(* IEC 61131-3 sources: plc-st-coding-agent/progress/evidence/f14_v10_full_20261113/jobs/custom_deepseek-v4pro (part 2) *)

(* ---- public-hard-02.raw_candidate_04.st ---- *)
(* ENGINEERING_CONTRACT
- Outputs conveyorLeft/deactivate in IDLE, PROCESSING and DONE; active only in MOVING state; no latch. PUB005.
- State machine: 0=IDLE waits sensor1 AND station1Start with valid length; 1=MOVING waits arrival at target sensor; 2=PROCESSING waits completion at current station 2..4; 3=DONE after station 5 arrival. PUB001/PUB002/PUB005.
- Movement direction: target station > current -> conveyorRight; target < current -> conveyorLeft; target == current stays at station for repeated processing step. PUB005.
- Completion signals are level-sensitive; on receiving completion, step advances, next sequence entry is queried, and movement restarts toward that station. PUB002.
- Final active sequence entry is station 5; arrival at 5 stops conveyor and enters DONE. A new start is permitted from DONE when the start condition is true. PUB003/PUB006.
- processLength validated 1..8; dynamic array indexing bounded by processLength; sequence values assumed to satisfy contract (2..4 processing, final 5). PUB004.
- Unspecified: exact restart behavior after DONE is level-sensitive on sensor1 and station1Start. No explicit reset input is used.
*)
(* CONTRACT_RULES [] *)
FUNCTION_BLOCK FlexibleProcessingControl
VAR_INPUT
    processLength : USINT;
    sensor1 : BOOL;
    sensor2 : BOOL;
    sensor3 : BOOL;
    sensor4 : BOOL;
    sensor5 : BOOL;
    station1Start : BOOL;
    station2Complete : BOOL;
    station3Complete : BOOL;
    station4Complete : BOOL;
    processSequence : ARRAY[1..8] OF USINT;
END_VAR
VAR_OUTPUT
    conveyorLeft : BOOL;
    conveyorRight : BOOL;
END_VAR
VAR
    local_state : USINT := 0; (* 0 = idle, 1 = moving, 2 = processing, 3 = done *)
    local_step : USINT := 0;
    local_target : USINT := 0;
    local_currentStation : USINT := 1;
    local_moveLeft : BOOL := FALSE;
    local_moveRight : BOOL := FALSE;
    local_arrival : BOOL := FALSE;
    local_complete : BOOL := FALSE;
END_VAR

(* Default outputs deactivated unless set by MOVING state *)
conveyorLeft := FALSE;
conveyorRight := FALSE;

CASE local_state OF
0: (* IDLE: wait for raw material at station 1 and start button *)
    IF processLength >= 1 AND processLength <= 8 AND sensor1 AND station1Start THEN
        local_step := 1;
        local_target := processSequence[1];
        local_currentStation := 1;
        IF local_target > local_currentStation THEN
            local_moveLeft := FALSE;
            local_moveRight := TRUE;
            conveyorLeft := FALSE;
            conveyorRight := TRUE;
            local_state := 1;
        ELSIF local_target < local_currentStation THEN
            local_moveLeft := TRUE;
            local_moveRight := FALSE;
            conveyorLeft := TRUE;
            conveyorRight := FALSE;
            local_state := 1;
        END_IF;
    END_IF;

1: (* MOVING: drive conveyor in chosen direction until target sensor detects arrival *)
    conveyorLeft := local_moveLeft;
    conveyorRight := local_moveRight;

    local_arrival := FALSE;
    IF local_target = 1 AND sensor1 THEN
        local_arrival := TRUE;
    ELSIF local_target = 2 AND sensor2 THEN
        local_arrival := TRUE;
    ELSIF local_target = 3 AND sensor3 THEN
        local_arrival := TRUE;
    ELSIF local_target = 4 AND sensor4 THEN
        local_arrival := TRUE;
    ELSIF local_target = 5 AND sensor5 THEN
        local_arrival := TRUE;
    END_IF;

    IF local_arrival THEN
        conveyorLeft := FALSE;
        conveyorRight := FALSE;
        local_moveLeft := FALSE;
        local_moveRight := FALSE;
        local_currentStation := local_target;

        IF local_currentStation = 5 THEN
            local_state := 3; (* final output station reached *)
        ELSE
            local_state := 2; (* processing station reached *)
        END_IF;
    END_IF;

2: (* PROCESSING: wait for completion signal at current processing station *)
    local_complete := FALSE;
    IF local_currentStation = 2 THEN
        local_complete := station2Complete;
    ELSIF local_currentStation = 3 THEN
        local_complete := station3Complete;
    ELSIF local_currentStation = 4 THEN
        local_complete := station4Complete;
    END_IF;

    IF local_complete THEN
        IF local_step < processLength THEN
            local_step := local_step + 1;
            local_target := processSequence[local_step];

            IF local_target > local_currentStation THEN
                local_moveLeft := FALSE;
                local_moveRight := TRUE;
                conveyorLeft := FALSE;
                conveyorRight := TRUE;
                local_state := 1;
            ELSIF local_target < local_currentStation THEN
                local_moveLeft := TRUE;
                local_moveRight := FALSE;
                conveyorLeft := TRUE;
                conveyorRight := FALSE;
                local_state := 1;
            ELSE
                (* Same station: remain in processing for the next sequence entry *)
                local_state := 2;
            END_IF;
        ELSE
            (* Invalid sequence: current processing station is not followed by final station 5 *)
            local_state := 3;
        END_IF;
    END_IF;

3: (* DONE: product delivered to station 5; optionally wait for next start *)
    IF processLength >= 1 AND processLength <= 8 AND sensor1 AND station1Start THEN
        local_step := 1;
        local_target := processSequence[1];
        local_currentStation := 1;
        IF local_target > local_currentStation THEN
            local_moveLeft := FALSE;
            local_moveRight := TRUE;
            conveyorLeft := FALSE;
            conveyorRight := TRUE;
            local_state := 1;
        ELSIF local_target < local_currentStation THEN
            local_moveLeft := TRUE;
            local_moveRight := FALSE;
            conveyorLeft := TRUE;
            conveyorRight := FALSE;
            local_state := 1;
        END_IF;
    END_IF;
END_CASE;

END_FUNCTION_BLOCK

(* ---- public-hard-03.candidate_01.st ---- *)
TYPE ST_Recipe :
STRUCT
    recipeID : INT;
    ingredientType : INT;
    ingredientRatio : REAL;
    productionTemperature : REAL;
END_STRUCT
END_TYPE;

FUNCTION_BLOCK FB_RecipeManagement
VAR_INPUT
    addRecipe : BOOL;
    deleteRecipe : BOOL;
    modifyRecipe : BOOL;
    queryRecipe : BOOL;
    recipeIn : ST_Recipe;
END_VAR
VAR_OUTPUT
    recipeAdded : BOOL;
    recipeDeleted : BOOL;
    recipeModified : BOOL;
    recipeQueryResult : ST_Recipe;
    error : BOOL;
    status : WORD;
END_VAR
VAR_IN_OUT
    recipe : ARRAY[1..10] OF ST_Recipe;
END_VAR
VAR
    tmp_i : INT;
    tmp_found : BOOL;
    tmp_index : INT;
    tmp_emptyIndex : INT;
    tmp_cmdCount : INT;
    tmp_emptyRecipe : ST_Recipe;
END_VAR

(*
ENGINEERING_CONTRACT
recipeAdded/Deleted/Modified: pulse TRUE only when exactly one matching request is TRUE and operation succeeds; not latched.
recipeQueryResult: valid only on successful query; otherwise zero struct. Not latched.
error/status: same-scan result; success/no command => error=FALSE,status=0. Error codes PUB003-PUB005, multiple commands => 16#8006.
recipe IN_OUT: caller retains; changed only on successful add/delete/modify. Add uses smallest empty index (PUB003).
Search ignores slots where recipeID=0. Units: raw REAL values; no scaling. Simultaneous commands are unsupported and modify nothing.
*)

(* CONTRACT_RULES [] *)

tmp_emptyRecipe.recipeID := 0;
tmp_emptyRecipe.ingredientType := 0;
tmp_emptyRecipe.ingredientRatio := 0.0;
tmp_emptyRecipe.productionTemperature := 0.0;

recipeAdded := FALSE;
recipeDeleted := FALSE;
recipeModified := FALSE;
recipeQueryResult := tmp_emptyRecipe;
error := FALSE;
status := 0;

tmp_cmdCount := 0;
IF addRecipe THEN
    tmp_cmdCount := tmp_cmdCount + 1;
END_IF;
IF deleteRecipe THEN
    tmp_cmdCount := tmp_cmdCount + 1;
END_IF;
IF modifyRecipe THEN
    tmp_cmdCount := tmp_cmdCount + 1;
END_IF;
IF queryRecipe THEN
    tmp_cmdCount := tmp_cmdCount + 1;
END_IF;

IF tmp_cmdCount > 1 THEN
    error := TRUE;
    status := 16#8006;
    RETURN;
END_IF;

IF addRecipe THEN
    tmp_found := FALSE;
    tmp_index := 0;
    FOR tmp_i := 1 TO 10 DO
        IF (recipe[tmp_i].recipeID <> 0) AND (recipe[tmp_i].recipeID = recipeIn.recipeID) THEN
            tmp_found := TRUE;
            tmp_index := tmp_i;
            EXIT;
        END_IF;
    END_FOR;

    IF tmp_found THEN
        error := TRUE;
        status := 16#8002;
    ELSE
        tmp_emptyIndex := 0;
        FOR tmp_i := 1 TO 10 DO
            IF recipe[tmp_i].recipeID = 0 THEN
                tmp_emptyIndex := tmp_i;
                EXIT;
            END_IF;
        END_FOR;

        IF tmp_emptyIndex = 0 THEN
            error := TRUE;
            status := 16#8003;
        ELSE
            recipe[tmp_emptyIndex] := recipeIn;
            recipeAdded := TRUE;
            error := FALSE;
            status := 0;
        END_IF;
    END_IF;
END_IF;

IF deleteRecipe THEN
    tmp_found := FALSE;
    tmp_index := 0;
    FOR tmp_i := 1 TO 10 DO
        IF (recipe[tmp_i].recipeID <> 0) AND (recipe[tmp_i].recipeID = recipeIn.recipeID) THEN
            tmp_found := TRUE;
            tmp_index := tmp_i;
            EXIT;
        END_IF;
    END_FOR;

    IF NOT tmp_found THEN
        error := TRUE;
        status := 16#8004;
    ELSE
        recipe[tmp_index] := tmp_emptyRecipe;
        recipeDeleted := TRUE;
        error := FALSE;
        status := 0;
    END_IF;
END_IF;

IF modifyRecipe THEN
    tmp_found := FALSE;
    tmp_index := 0;
    FOR tmp_i := 1 TO 10 DO
        IF (recipe[tmp_i].recipeID <> 0) AND (recipe[tmp_i].recipeID = recipeIn.recipeID) THEN
            tmp_found := TRUE;
            tmp_index := tmp_i;
            EXIT;
        END_IF;
    END_FOR;

    IF NOT tmp_found THEN
        error := TRUE;
        status := 16#8005;
    ELSE
        recipe[tmp_index] := recipeIn;
        recipeModified := TRUE;
        error := FALSE;
        status := 0;
    END_IF;
END_IF;

IF queryRecipe THEN
    tmp_found := FALSE;
    tmp_index := 0;
    FOR tmp_i := 1 TO 10 DO
        IF (recipe[tmp_i].recipeID <> 0) AND (recipe[tmp_i].recipeID = recipeIn.recipeID) THEN
            tmp_found := TRUE;
            tmp_index := tmp_i;
            EXIT;
        END_IF;
    END_FOR;

    IF NOT tmp_found THEN
        error := TRUE;
        status := 16#8001;
    ELSE
        recipeQueryResult := recipe[tmp_index];
        error := FALSE;
        status := 0;
    END_IF;
END_IF;

END_FUNCTION_BLOCK

(* ---- public-hard-03.candidate_02.st ---- *)
TYPE ST_Recipe :
STRUCT
    recipeID : INT;
    ingredientType : INT;
    ingredientRatio : REAL;
    productionTemperature : REAL;
END_STRUCT
END_TYPE;

FUNCTION_BLOCK FB_RecipeManagement
VAR_INPUT
    addRecipe : BOOL;
    deleteRecipe : BOOL;
    modifyRecipe : BOOL;
    queryRecipe : BOOL;
    recipeIn : ST_Recipe;
END_VAR
VAR_OUTPUT
    recipeAdded : BOOL;
    recipeDeleted : BOOL;
    recipeModified : BOOL;
    recipeQueryResult : ST_Recipe;
    error : BOOL;
    status : WORD;
END_VAR
VAR_IN_OUT
    recipe : ARRAY[1..10] OF ST_Recipe;
END_VAR
VAR
    tmp_i : INT;
    tmp_found : BOOL;
    tmp_index : INT;
    tmp_emptyIndex : INT;
    tmp_cmdCount : INT;
    tmp_emptyRecipe : ST_Recipe;
    tmp_addReq : BOOL;
    tmp_deleteReq : BOOL;
    tmp_modifyReq : BOOL;
    tmp_queryReq : BOOL;
    prevAdd : BOOL := FALSE;
    prevDelete : BOOL := FALSE;
    prevModify : BOOL := FALSE;
    prevQuery : BOOL := FALSE;
END_VAR

(*
ENGINEERING_CONTRACT
Request signals are edge-triggered (rising edge only).
recipeAdded/Deleted/Modified: one-scan pulse on successful operation; otherwise FALSE.
recipeQueryResult: valid only in the scan of a successful query; zero struct otherwise.
error/status: same-scan result; success/no edge => error=FALSE,status=0.
Simultaneous rising command edges => error=TRUE,status=16#8006; database unchanged.
Database in recipe[] retains state between scans; add uses smallest empty index.
*)

(* CONTRACT_RULES [] *)

tmp_emptyRecipe.recipeID := 0;
tmp_emptyRecipe.ingredientType := 0;
tmp_emptyRecipe.ingredientRatio := 0.0;
tmp_emptyRecipe.productionTemperature := 0.0;

recipeAdded := FALSE;
recipeDeleted := FALSE;
recipeModified := FALSE;
recipeQueryResult := tmp_emptyRecipe;
error := FALSE;
status := 0;

tmp_addReq := addRecipe AND NOT prevAdd;
tmp_deleteReq := deleteRecipe AND NOT prevDelete;
tmp_modifyReq := modifyRecipe AND NOT prevModify;
tmp_queryReq := queryRecipe AND NOT prevQuery;

prevAdd := addRecipe;
prevDelete := deleteRecipe;
prevModify := modifyRecipe;
prevQuery := queryRecipe;

tmp_cmdCount := 0;
IF tmp_addReq THEN
    tmp_cmdCount := tmp_cmdCount + 1;
END_IF;
IF tmp_deleteReq THEN
    tmp_cmdCount := tmp_cmdCount + 1;
END_IF;
IF tmp_modifyReq THEN
    tmp_cmdCount := tmp_cmdCount + 1;
END_IF;
IF tmp_queryReq THEN
    tmp_cmdCount := tmp_cmdCount + 1;
END_IF;

IF tmp_cmdCount > 1 THEN
    error := TRUE;
    status := 16#8006;
    RETURN;
END_IF;

IF tmp_addReq THEN
    tmp_found := FALSE;
    tmp_index := 0;
    FOR tmp_i := 1 TO 10 DO
        IF (recipe[tmp_i].recipeID <> 0) AND (recipe[tmp_i].recipeID = recipeIn.recipeID) THEN
            tmp_found := TRUE;
            tmp_index := tmp_i;
            EXIT;
        END_IF;
    END_FOR;

    IF tmp_found THEN
        error := TRUE;
        status := 16#8002;
    ELSE
        tmp_emptyIndex := 0;
        FOR tmp_i := 1 TO 10 DO
            IF recipe[tmp_i].recipeID = 0 THEN
                tmp_emptyIndex := tmp_i;
                EXIT;
            END_IF;
        END_FOR;

        IF tmp_emptyIndex = 0 THEN
            error := TRUE;
            status := 16#8003;
        ELSE
            recipe[tmp_emptyIndex] := recipeIn;
            recipeAdded := TRUE;
            error := FALSE;
            status := 0;
        END_IF;
    END_IF;
END_IF;

IF tmp_deleteReq THEN
    tmp_found := FALSE;
    tmp_index := 0;
    FOR tmp_i := 1 TO 10 DO
        IF (recipe[tmp_i].recipeID <> 0) AND (recipe[tmp_i].recipeID = recipeIn.recipeID) THEN
            tmp_found := TRUE;
            tmp_index := tmp_i;
            EXIT;
        END_IF;
    END_FOR;

    IF NOT tmp_found THEN
        error := TRUE;
        status := 16#8004;
    ELSE
        recipe[tmp_index] := tmp_emptyRecipe;
        recipeDeleted := TRUE;
        error := FALSE;
        status := 0;
    END_IF;
END_IF;

IF tmp_modifyReq THEN
    tmp_found := FALSE;
    tmp_index := 0;
    FOR tmp_i := 1 TO 10 DO
        IF (recipe[tmp_i].recipeID <> 0) AND (recipe[tmp_i].recipeID = recipeIn.recipeID) THEN
            tmp_found := TRUE;
            tmp_index := tmp_i;
            EXIT;
        END_IF;
    END_FOR;

    IF NOT tmp_found THEN
        error := TRUE;
        status := 16#8005;
    ELSE
        recipe[tmp_index] := recipeIn;
        recipeModified := TRUE;
        error := FALSE;
        status := 0;
    END_IF;
END_IF;

IF tmp_queryReq THEN
    tmp_found := FALSE;
    tmp_index := 0;
    FOR tmp_i := 1 TO 10 DO
        IF (recipe[tmp_i].recipeID <> 0) AND (recipe[tmp_i].recipeID = recipeIn.recipeID) THEN
            tmp_found := TRUE;
            tmp_index := tmp_i;
            EXIT;
        END_IF;
    END_FOR;

    IF NOT tmp_found THEN
        error := TRUE;
        status := 16#8001;
    ELSE
        recipeQueryResult := recipe[tmp_index];
        error := FALSE;
        status := 0;
    END_IF;
END_IF;

END_FUNCTION_BLOCK

(* ---- public-hard-03.candidate_03.st ---- *)
TYPE ST_Recipe :
STRUCT
    recipeID : INT;
    ingredientType : INT;
    ingredientRatio : REAL;
    productionTemperature : REAL;
END_STRUCT
END_TYPE;

FUNCTION_BLOCK FB_RecipeManagement
VAR_INPUT
    addRecipe : BOOL;
    deleteRecipe : BOOL;
    modifyRecipe : BOOL;
    queryRecipe : BOOL;
    recipeIn : ST_Recipe;
END_VAR
VAR_OUTPUT
    recipeAdded : BOOL;
    recipeDeleted : BOOL;
    recipeModified : BOOL;
    recipeQueryResult : ST_Recipe;
    error : BOOL;
    status : WORD;
END_VAR
VAR_IN_OUT
    recipe : ARRAY[1..10] OF ST_Recipe;
END_VAR
VAR
    tmp_i : INT;
    tmp_found : BOOL;
    tmp_index : INT;
    tmp_emptyIndex : INT;
    tmp_emptyRecipe : ST_Recipe;
END_VAR

(*
ENGINEERING_CONTRACT
recipeAdded/Deleted/Modified: pulse TRUE only when corresponding request is TRUE and operation succeeds; not latched.
recipeQueryResult: valid only on successful query; otherwise zero struct. Not latched.
error/status: same-scan result; success/no command => error=FALSE,status=0.
Search ignores slots where recipeID=0. Units: raw REAL values; no scaling.
Simultaneous commands are not specified by the public contract; implementation processes all active commands in the
present scan using the defined operation order add, delete, modify, query. No extra priority or 8006 code is invented.
*)

(* CONTRACT_RULES [] *)

tmp_emptyRecipe.recipeID := 0;
tmp_emptyRecipe.ingredientType := 0;
tmp_emptyRecipe.ingredientRatio := 0.0;
tmp_emptyRecipe.productionTemperature := 0.0;

recipeAdded := FALSE;
recipeDeleted := FALSE;
recipeModified := FALSE;
recipeQueryResult := tmp_emptyRecipe;
error := FALSE;
status := 0;

IF addRecipe THEN
    tmp_found := FALSE;
    tmp_index := 0;
    FOR tmp_i := 1 TO 10 DO
        IF (recipe[tmp_i].recipeID <> 0) AND (recipe[tmp_i].recipeID = recipeIn.recipeID) THEN
            tmp_found := TRUE;
            tmp_index := tmp_i;
            EXIT;
        END_IF;
    END_FOR;

    IF tmp_found THEN
        error := TRUE;
        status := 16#8002;
    ELSE
        tmp_emptyIndex := 0;
        FOR tmp_i := 1 TO 10 DO
            IF recipe[tmp_i].recipeID = 0 THEN
                tmp_emptyIndex := tmp_i;
                EXIT;
            END_IF;
        END_FOR;

        IF tmp_emptyIndex = 0 THEN
            error := TRUE;
            status := 16#8003;
        ELSE
            recipe[tmp_emptyIndex] := recipeIn;
            recipeAdded := TRUE;
            error := FALSE;
            status := 0;
        END_IF;
    END_IF;
END_IF;

IF deleteRecipe THEN
    tmp_found := FALSE;
    tmp_index := 0;
    FOR tmp_i := 1 TO 10 DO
        IF (recipe[tmp_i].recipeID <> 0) AND (recipe[tmp_i].recipeID = recipeIn.recipeID) THEN
            tmp_found := TRUE;
            tmp_index := tmp_i;
            EXIT;
        END_IF;
    END_FOR;

    IF NOT tmp_found THEN
        error := TRUE;
        status := 16#8004;
    ELSE
        recipe[tmp_index] := tmp_emptyRecipe;
        recipeDeleted := TRUE;
        error := FALSE;
        status := 0;
    END_IF;
END_IF;

IF modifyRecipe THEN
    tmp_found := FALSE;
    tmp_index := 0;
    FOR tmp_i := 1 TO 10 DO
        IF (recipe[tmp_i].recipeID <> 0) AND (recipe[tmp_i].recipeID = recipeIn.recipeID) THEN
            tmp_found := TRUE;
            tmp_index := tmp_i;
            EXIT;
        END_IF;
    END_FOR;

    IF NOT tmp_found THEN
        error := TRUE;
        status := 16#8005;
    ELSE
        recipe[tmp_index] := recipeIn;
        recipeModified := TRUE;
        error := FALSE;
        status := 0;
    END_IF;
END_IF;

IF queryRecipe THEN
    tmp_found := FALSE;
    tmp_index := 0;
    FOR tmp_i := 1 TO 10 DO
        IF (recipe[tmp_i].recipeID <> 0) AND (recipe[tmp_i].recipeID = recipeIn.recipeID) THEN
            tmp_found := TRUE;
            tmp_index := tmp_i;
            EXIT;
        END_IF;
    END_FOR;

    IF NOT tmp_found THEN
        error := TRUE;
        status := 16#8001;
    ELSE
        recipeQueryResult := recipe[tmp_index];
        error := FALSE;
        status := 0;
    END_IF;
END_IF;

END_FUNCTION_BLOCK

(* ---- public-hard-03.candidate_04.st ---- *)
TYPE ST_Recipe :
STRUCT
    recipeID : INT;
    ingredientType : INT;
    ingredientRatio : REAL;
    productionTemperature : REAL;
END_STRUCT
END_TYPE;

FUNCTION_BLOCK FB_RecipeManagement
VAR_INPUT
    addRecipe : BOOL;
    deleteRecipe : BOOL;
    modifyRecipe : BOOL;
    queryRecipe : BOOL;
    recipeIn : ST_Recipe;
END_VAR
VAR_OUTPUT
    recipeAdded : BOOL;
    recipeDeleted : BOOL;
    recipeModified : BOOL;
    recipeQueryResult : ST_Recipe;
    error : BOOL;
    status : WORD;
END_VAR
VAR_IN_OUT
    recipe : ARRAY[1..10] OF ST_Recipe;
END_VAR
VAR
    tmp_i : INT;
    tmp_found : BOOL;
    tmp_index : INT;
    tmp_emptyIndex : INT;
    tmp_cmdCount : INT;
    tmp_emptyRecipe : ST_Recipe;
END_VAR

(*
ENGINEERING_CONTRACT
recipeAdded/Deleted/Modified: pulse TRUE only when exactly one matching request is TRUE and operation succeeds; not latched.
recipeQueryResult: valid only on successful query; otherwise zero struct. Not latched.
error/status: same-scan result; success/no command => error=FALSE,status=0. Error codes PUB003-PUB005, multiple commands => 16#8006.
recipe IN_OUT: caller retains; changed only on successful add/delete/modify. Add uses smallest empty index (PUB003).
Search ignores slots where recipeID=0 for query/delete/modify. Add treats recipeIn.recipeID=0 as reserved/invalid and never stores it.
Units: raw REAL values; no scaling. Simultaneous commands are unsupported and modify nothing.
*)

(* CONTRACT_RULES [] *)

tmp_emptyRecipe.recipeID := 0;
tmp_emptyRecipe.ingredientType := 0;
tmp_emptyRecipe.ingredientRatio := 0.0;
tmp_emptyRecipe.productionTemperature := 0.0;

recipeAdded := FALSE;
recipeDeleted := FALSE;
recipeModified := FALSE;
recipeQueryResult := tmp_emptyRecipe;
error := FALSE;
status := 0;

tmp_cmdCount := 0;
IF addRecipe THEN
    tmp_cmdCount := tmp_cmdCount + 1;
END_IF;
IF deleteRecipe THEN
    tmp_cmdCount := tmp_cmdCount + 1;
END_IF;
IF modifyRecipe THEN
    tmp_cmdCount := tmp_cmdCount + 1;
END_IF;
IF queryRecipe THEN
    tmp_cmdCount := tmp_cmdCount + 1;
END_IF;

IF tmp_cmdCount > 1 THEN
    error := TRUE;
    status := 16#8006;
    RETURN;
END_IF;

IF addRecipe THEN
    tmp_found := FALSE;
    tmp_index := 0;
    FOR tmp_i := 1 TO 10 DO
        IF recipe[tmp_i].recipeID = recipeIn.recipeID THEN
            tmp_found := TRUE;
            tmp_index := tmp_i;
            EXIT;
        END_IF;
    END_FOR;

    IF tmp_found THEN
        error := TRUE;
        status := 16#8002;
    ELSE
        tmp_emptyIndex := 0;
        FOR tmp_i := 1 TO 10 DO
            IF recipe[tmp_i].recipeID = 0 THEN
                tmp_emptyIndex := tmp_i;
                EXIT;
            END_IF;
        END_FOR;

        IF tmp_emptyIndex = 0 THEN
            error := TRUE;
            status := 16#8003;
        ELSE
            recipe[tmp_emptyIndex] := recipeIn;
            recipeAdded := TRUE;
            error := FALSE;
            status := 0;
        END_IF;
    END_IF;
END_IF;

IF deleteRecipe THEN
    tmp_found := FALSE;
    tmp_index := 0;
    FOR tmp_i := 1 TO 10 DO
        IF (recipe[tmp_i].recipeID <> 0) AND (recipe[tmp_i].recipeID = recipeIn.recipeID) THEN
            tmp_found := TRUE;
            tmp_index := tmp_i;
            EXIT;
        END_IF;
    END_FOR;

    IF NOT tmp_found THEN
        error := TRUE;
        status := 16#8004;
    ELSE
        recipe[tmp_index] := tmp_emptyRecipe;
        recipeDeleted := TRUE;
        error := FALSE;
        status := 0;
    END_IF;
END_IF;

IF modifyRecipe THEN
    tmp_found := FALSE;
    tmp_index := 0;
    FOR tmp_i := 1 TO 10 DO
        IF (recipe[tmp_i].recipeID <> 0) AND (recipe[tmp_i].recipeID = recipeIn.recipeID) THEN
            tmp_found := TRUE;
            tmp_index := tmp_i;
            EXIT;
        END_IF;
    END_FOR;

    IF NOT tmp_found THEN
        error := TRUE;
        status := 16#8005;
    ELSE
        recipe[tmp_index] := recipeIn;
        recipeModified := TRUE;
        error := FALSE;
        status := 0;
    END_IF;
END_IF;

IF queryRecipe THEN
    tmp_found := FALSE;
    tmp_index := 0;
    FOR tmp_i := 1 TO 10 DO
        IF (recipe[tmp_i].recipeID <> 0) AND (recipe[tmp_i].recipeID = recipeIn.recipeID) THEN
            tmp_found := TRUE;
            tmp_index := tmp_i;
            EXIT;
        END_IF;
    END_FOR;

    IF NOT tmp_found THEN
        error := TRUE;
        status := 16#8001;
    ELSE
        recipeQueryResult := recipe[tmp_index];
        error := FALSE;
        status := 0;
    END_IF;
END_IF;

END_FUNCTION_BLOCK

(* ---- public-hard-03.raw_candidate_01.st ---- *)
TYPE ST_Recipe :
STRUCT
    recipeID : INT;
    ingredientType : INT;
    ingredientRatio : REAL;
    productionTemperature : REAL;
END_STRUCT
END_TYPE

FUNCTION_BLOCK FB_RecipeManagement
VAR_INPUT
    addRecipe : BOOL;
    deleteRecipe : BOOL;
    modifyRecipe : BOOL;
    queryRecipe : BOOL;
    recipeIn : ST_Recipe;
END_VAR
VAR_OUTPUT
    recipeAdded : BOOL;
    recipeDeleted : BOOL;
    recipeModified : BOOL;
    recipeQueryResult : ST_Recipe;
    error : BOOL;
    status : WORD;
END_VAR
VAR_IN_OUT
    recipe : ARRAY[1..10] OF ST_Recipe;
END_VAR
VAR
    tmp_i : INT;
    tmp_found : BOOL;
    tmp_index : INT;
    tmp_emptyIndex : INT;
    tmp_cmdCount : INT;
    tmp_emptyRecipe : ST_Recipe;
END_VAR

(*
ENGINEERING_CONTRACT
recipeAdded/Deleted/Modified: pulse TRUE only when exactly one matching request is TRUE and operation succeeds; not latched.
recipeQueryResult: valid only on successful query; otherwise zero struct. Not latched.
error/status: same-scan result; success/no command => error=FALSE,status=0. Error codes PUB003-PUB005, multiple commands => 16#8006.
recipe IN_OUT: caller retains; changed only on successful add/delete/modify. Add uses smallest empty index (PUB003).
Search ignores slots where recipeID=0. Units: raw REAL values; no scaling. Simultaneous commands are unsupported and modify nothing.
*)

(* CONTRACT_RULES [] *)

tmp_emptyRecipe.recipeID := 0;
tmp_emptyRecipe.ingredientType := 0;
tmp_emptyRecipe.ingredientRatio := 0.0;
tmp_emptyRecipe.productionTemperature := 0.0;

recipeAdded := FALSE;
recipeDeleted := FALSE;
recipeModified := FALSE;
recipeQueryResult := tmp_emptyRecipe;
error := FALSE;
status := 0;

tmp_cmdCount := 0;
IF addRecipe THEN
    tmp_cmdCount := tmp_cmdCount + 1;
END_IF;
IF deleteRecipe THEN
    tmp_cmdCount := tmp_cmdCount + 1;
END_IF;
IF modifyRecipe THEN
    tmp_cmdCount := tmp_cmdCount + 1;
END_IF;
IF queryRecipe THEN
    tmp_cmdCount := tmp_cmdCount + 1;
END_IF;

IF tmp_cmdCount > 1 THEN
    error := TRUE;
    status := 16#8006;
    RETURN;
END_IF;

IF addRecipe THEN
    tmp_found := FALSE;
    tmp_index := 0;
    FOR tmp_i := 1 TO 10 DO
        IF (recipe[tmp_i].recipeID <> 0) AND (recipe[tmp_i].recipeID = recipeIn.recipeID) THEN
            tmp_found := TRUE;
            tmp_index := tmp_i;
            EXIT;
        END_IF;
    END_FOR;

    IF tmp_found THEN
        error := TRUE;
        status := 16#8002;
    ELSE
        tmp_emptyIndex := 0;
        FOR tmp_i := 1 TO 10 DO
            IF recipe[tmp_i].recipeID = 0 THEN
                tmp_emptyIndex := tmp_i;
                EXIT;
            END_IF;
        END_FOR;

        IF tmp_emptyIndex = 0 THEN
            error := TRUE;
            status := 16#8003;
        ELSE
            recipe[tmp_emptyIndex] := recipeIn;
            recipeAdded := TRUE;
            error := FALSE;
            status := 0;
        END_IF;
    END_IF;
END_IF;

IF deleteRecipe THEN
    tmp_found := FALSE;
    tmp_index := 0;
    FOR tmp_i := 1 TO 10 DO
        IF (recipe[tmp_i].recipeID <> 0) AND (recipe[tmp_i].recipeID = recipeIn.recipeID) THEN
            tmp_found := TRUE;
            tmp_index := tmp_i;
            EXIT;
        END_IF;
    END_FOR;

    IF NOT tmp_found THEN
        error := TRUE;
        status := 16#8004;
    ELSE
        recipe[tmp_index] := tmp_emptyRecipe;
        recipeDeleted := TRUE;
        error := FALSE;
        status := 0;
    END_IF;
END_IF;

IF modifyRecipe THEN
    tmp_found := FALSE;
    tmp_index := 0;
    FOR tmp_i := 1 TO 10 DO
        IF (recipe[tmp_i].recipeID <> 0) AND (recipe[tmp_i].recipeID = recipeIn.recipeID) THEN
            tmp_found := TRUE;
            tmp_index := tmp_i;
            EXIT;
        END_IF;
    END_FOR;

    IF NOT tmp_found THEN
        error := TRUE;
        status := 16#8005;
    ELSE
        recipe[tmp_index] := recipeIn;
        recipeModified := TRUE;
        error := FALSE;
        status := 0;
    END_IF;
END_IF;

IF queryRecipe THEN
    tmp_found := FALSE;
    tmp_index := 0;
    FOR tmp_i := 1 TO 10 DO
        IF (recipe[tmp_i].recipeID <> 0) AND (recipe[tmp_i].recipeID = recipeIn.recipeID) THEN
            tmp_found := TRUE;
            tmp_index := tmp_i;
            EXIT;
        END_IF;
    END_FOR;

    IF NOT tmp_found THEN
        error := TRUE;
        status := 16#8001;
    ELSE
        recipeQueryResult := recipe[tmp_index];
        error := FALSE;
        status := 0;
    END_IF;
END_IF;

END_FUNCTION_BLOCK

(* ---- public-hard-03.raw_candidate_02.st ---- *)
TYPE ST_Recipe :
STRUCT
    recipeID : INT;
    ingredientType : INT;
    ingredientRatio : REAL;
    productionTemperature : REAL;
END_STRUCT
END_TYPE;

FUNCTION_BLOCK FB_RecipeManagement
VAR_INPUT
    addRecipe : BOOL;
    deleteRecipe : BOOL;
    modifyRecipe : BOOL;
    queryRecipe : BOOL;
    recipeIn : ST_Recipe;
END_VAR
VAR_OUTPUT
    recipeAdded : BOOL;
    recipeDeleted : BOOL;
    recipeModified : BOOL;
    recipeQueryResult : ST_Recipe;
    error : BOOL;
    status : WORD;
END_VAR
VAR_IN_OUT
    recipe : ARRAY[1..10] OF ST_Recipe;
END_VAR
VAR
    tmp_i : INT;
    tmp_found : BOOL;
    tmp_index : INT;
    tmp_emptyIndex : INT;
    tmp_cmdCount : INT;
    tmp_emptyRecipe : ST_Recipe;
    tmp_addReq : BOOL;
    tmp_deleteReq : BOOL;
    tmp_modifyReq : BOOL;
    tmp_queryReq : BOOL;
    prevAdd : BOOL := FALSE;
    prevDelete : BOOL := FALSE;
    prevModify : BOOL := FALSE;
    prevQuery : BOOL := FALSE;
END_VAR

(*
ENGINEERING_CONTRACT
Request signals are edge-triggered (rising edge only).
recipeAdded/Deleted/Modified: one-scan pulse on successful operation; otherwise FALSE.
recipeQueryResult: valid only in the scan of a successful query; zero struct otherwise.
error/status: same-scan result; success/no edge => error=FALSE,status=0.
Simultaneous rising command edges => error=TRUE,status=16#8006; database unchanged.
Database in recipe[] retains state between scans; add uses smallest empty index.
*)

(* CONTRACT_RULES [] *)

tmp_emptyRecipe.recipeID := 0;
tmp_emptyRecipe.ingredientType := 0;
tmp_emptyRecipe.ingredientRatio := 0.0;
tmp_emptyRecipe.productionTemperature := 0.0;

recipeAdded := FALSE;
recipeDeleted := FALSE;
recipeModified := FALSE;
recipeQueryResult := tmp_emptyRecipe;
error := FALSE;
status := 0;

tmp_addReq := addRecipe AND NOT prevAdd;
tmp_deleteReq := deleteRecipe AND NOT prevDelete;
tmp_modifyReq := modifyRecipe AND NOT prevModify;
tmp_queryReq := queryRecipe AND NOT prevQuery;

prevAdd := addRecipe;
prevDelete := deleteRecipe;
prevModify := modifyRecipe;
prevQuery := queryRecipe;

tmp_cmdCount := 0;
IF tmp_addReq THEN
    tmp_cmdCount := tmp_cmdCount + 1;
END_IF;
IF tmp_deleteReq THEN
    tmp_cmdCount := tmp_cmdCount + 1;
END_IF;
IF tmp_modifyReq THEN
    tmp_cmdCount := tmp_cmdCount + 1;
END_IF;
IF tmp_queryReq THEN
    tmp_cmdCount := tmp_cmdCount + 1;
END_IF;

IF tmp_cmdCount > 1 THEN
    error := TRUE;
    status := 16#8006;
    RETURN;
END_IF;

IF tmp_addReq THEN
    tmp_found := FALSE;
    tmp_index := 0;
    FOR tmp_i := 1 TO 10 DO
        IF (recipe[tmp_i].recipeID <> 0) AND (recipe[tmp_i].recipeID = recipeIn.recipeID) THEN
            tmp_found := TRUE;
            tmp_index := tmp_i;
            EXIT;
        END_IF;
    END_FOR;

    IF tmp_found THEN
        error := TRUE;
        status := 16#8002;
    ELSE
        tmp_emptyIndex := 0;
        FOR tmp_i := 1 TO 10 DO
            IF recipe[tmp_i].recipeID = 0 THEN
                tmp_emptyIndex := tmp_i;
                EXIT;
            END_IF;
        END_FOR;

        IF tmp_emptyIndex = 0 THEN
            error := TRUE;
            status := 16#8003;
        ELSE
            recipe[tmp_emptyIndex] := recipeIn;
            recipeAdded := TRUE;
            error := FALSE;
            status := 0;
        END_IF;
    END_IF;
END_IF;

IF tmp_deleteReq THEN
    tmp_found := FALSE;
    tmp_index := 0;
    FOR tmp_i := 1 TO 10 DO
        IF (recipe[tmp_i].recipeID <> 0) AND (recipe[tmp_i].recipeID = recipeIn.recipeID) THEN
            tmp_found := TRUE;
            tmp_index := tmp_i;
            EXIT;
        END_IF;
    END_FOR;

    IF NOT tmp_found THEN
        error := TRUE;
        status := 16#8004;
    ELSE
        recipe[tmp_index] := tmp_emptyRecipe;
        recipeDeleted := TRUE;
        error := FALSE;
        status := 0;
    END_IF;
END_IF;

IF tmp_modifyReq THEN
    tmp_found := FALSE;
    tmp_index := 0;
    FOR tmp_i := 1 TO 10 DO
        IF (recipe[tmp_i].recipeID <> 0) AND (recipe[tmp_i].recipeID = recipeIn.recipeID) THEN
            tmp_found := TRUE;
            tmp_index := tmp_i;
            EXIT;
        END_IF;
    END_FOR;

    IF NOT tmp_found THEN
        error := TRUE;
        status := 16#8005;
    ELSE
        recipe[tmp_index] := recipeIn;
        recipeModified := TRUE;
        error := FALSE;
        status := 0;
    END_IF;
END_IF;

IF tmp_queryReq THEN
    tmp_found := FALSE;
    tmp_index := 0;
    FOR tmp_i := 1 TO 10 DO
        IF (recipe[tmp_i].recipeID <> 0) AND (recipe[tmp_i].recipeID = recipeIn.recipeID) THEN
            tmp_found := TRUE;
            tmp_index := tmp_i;
            EXIT;
        END_IF;
    END_FOR;

    IF NOT tmp_found THEN
        error := TRUE;
        status := 16#8001;
    ELSE
        recipeQueryResult := recipe[tmp_index];
        error := FALSE;
        status := 0;
    END_IF;
END_IF;

END_FUNCTION_BLOCK

(* ---- public-hard-03.raw_candidate_03.st ---- *)
TYPE ST_Recipe :
STRUCT
    recipeID : INT;
    ingredientType : INT;
    ingredientRatio : REAL;
    productionTemperature : REAL;
END_STRUCT
END_TYPE;

FUNCTION_BLOCK FB_RecipeManagement
VAR_INPUT
    addRecipe : BOOL;
    deleteRecipe : BOOL;
    modifyRecipe : BOOL;
    queryRecipe : BOOL;
    recipeIn : ST_Recipe;
END_VAR
VAR_OUTPUT
    recipeAdded : BOOL;
    recipeDeleted : BOOL;
    recipeModified : BOOL;
    recipeQueryResult : ST_Recipe;
    error : BOOL;
    status : WORD;
END_VAR
VAR_IN_OUT
    recipe : ARRAY[1..10] OF ST_Recipe;
END_VAR
VAR
    tmp_i : INT;
    tmp_found : BOOL;
    tmp_index : INT;
    tmp_emptyIndex : INT;
    tmp_emptyRecipe : ST_Recipe;
END_VAR

(*
ENGINEERING_CONTRACT
recipeAdded/Deleted/Modified: pulse TRUE only when corresponding request is TRUE and operation succeeds; not latched.
recipeQueryResult: valid only on successful query; otherwise zero struct. Not latched.
error/status: same-scan result; success/no command => error=FALSE,status=0.
Search ignores slots where recipeID=0. Units: raw REAL values; no scaling.
Simultaneous commands are not specified by the public contract; implementation processes all active commands in the
present scan using the defined operation order add, delete, modify, query. No extra priority or 8006 code is invented.
*)

(* CONTRACT_RULES [] *)

tmp_emptyRecipe.recipeID := 0;
tmp_emptyRecipe.ingredientType := 0;
tmp_emptyRecipe.ingredientRatio := 0.0;
tmp_emptyRecipe.productionTemperature := 0.0;

recipeAdded := FALSE;
recipeDeleted := FALSE;
recipeModified := FALSE;
recipeQueryResult := tmp_emptyRecipe;
error := FALSE;
status := 0;

IF addRecipe THEN
    tmp_found := FALSE;
    tmp_index := 0;
    FOR tmp_i := 1 TO 10 DO
        IF (recipe[tmp_i].recipeID <> 0) AND (recipe[tmp_i].recipeID = recipeIn.recipeID) THEN
            tmp_found := TRUE;
            tmp_index := tmp_i;
            EXIT;
        END_IF;
    END_FOR;

    IF tmp_found THEN
        error := TRUE;
        status := 16#8002;
    ELSE
        tmp_emptyIndex := 0;
        FOR tmp_i := 1 TO 10 DO
            IF recipe[tmp_i].recipeID = 0 THEN
                tmp_emptyIndex := tmp_i;
                EXIT;
            END_IF;
        END_FOR;

        IF tmp_emptyIndex = 0 THEN
            error := TRUE;
            status := 16#8003;
        ELSE
            recipe[tmp_emptyIndex] := recipeIn;
            recipeAdded := TRUE;
            error := FALSE;
            status := 0;
        END_IF;
    END_IF;
END_IF;

IF deleteRecipe THEN
    tmp_found := FALSE;
    tmp_index := 0;
    FOR tmp_i := 1 TO 10 DO
        IF (recipe[tmp_i].recipeID <> 0) AND (recipe[tmp_i].recipeID = recipeIn.recipeID) THEN
            tmp_found := TRUE;
            tmp_index := tmp_i;
            EXIT;
        END_IF;
    END_FOR;

    IF NOT tmp_found THEN
        error := TRUE;
        status := 16#8004;
    ELSE
        recipe[tmp_index] := tmp_emptyRecipe;
        recipeDeleted := TRUE;
        error := FALSE;
        status := 0;
    END_IF;
END_IF;

IF modifyRecipe THEN
    tmp_found := FALSE;
    tmp_index := 0;
    FOR tmp_i := 1 TO 10 DO
        IF (recipe[tmp_i].recipeID <> 0) AND (recipe[tmp_i].recipeID = recipeIn.recipeID) THEN
            tmp_found := TRUE;
            tmp_index := tmp_i;
            EXIT;
        END_IF;
    END_FOR;

    IF NOT tmp_found THEN
        error := TRUE;
        status := 16#8005;
    ELSE
        recipe[tmp_index] := recipeIn;
        recipeModified := TRUE;
        error := FALSE;
        status := 0;
    END_IF;
END_IF;

IF queryRecipe THEN
    tmp_found := FALSE;
    tmp_index := 0;
    FOR tmp_i := 1 TO 10 DO
        IF (recipe[tmp_i].recipeID <> 0) AND (recipe[tmp_i].recipeID = recipeIn.recipeID) THEN
            tmp_found := TRUE;
            tmp_index := tmp_i;
            EXIT;
        END_IF;
    END_FOR;

    IF NOT tmp_found THEN
        error := TRUE;
        status := 16#8001;
    ELSE
        recipeQueryResult := recipe[tmp_index];
        error := FALSE;
        status := 0;
    END_IF;
END_IF;

END_FUNCTION_BLOCK

(* ---- public-hard-03.raw_candidate_04.st ---- *)
TYPE ST_Recipe :
STRUCT
    recipeID : INT;
    ingredientType : INT;
    ingredientRatio : REAL;
    productionTemperature : REAL;
END_STRUCT
END_TYPE;

FUNCTION_BLOCK FB_RecipeManagement
VAR_INPUT
    addRecipe : BOOL;
    deleteRecipe : BOOL;
    modifyRecipe : BOOL;
    queryRecipe : BOOL;
    recipeIn : ST_Recipe;
END_VAR
VAR_OUTPUT
    recipeAdded : BOOL;
    recipeDeleted : BOOL;
    recipeModified : BOOL;
    recipeQueryResult : ST_Recipe;
    error : BOOL;
    status : WORD;
END_VAR
VAR_IN_OUT
    recipe : ARRAY[1..10] OF ST_Recipe;
END_VAR
VAR
    tmp_i : INT;
    tmp_found : BOOL;
    tmp_index : INT;
    tmp_emptyIndex : INT;
    tmp_cmdCount : INT;
    tmp_emptyRecipe : ST_Recipe;
END_VAR

(*
ENGINEERING_CONTRACT
recipeAdded/Deleted/Modified: pulse TRUE only when exactly one matching request is TRUE and operation succeeds; not latched.
recipeQueryResult: valid only on successful query; otherwise zero struct. Not latched.
error/status: same-scan result; success/no command => error=FALSE,status=0. Error codes PUB003-PUB005, multiple commands => 16#8006.
recipe IN_OUT: caller retains; changed only on successful add/delete/modify. Add uses smallest empty index (PUB003).
Search ignores slots where recipeID=0 for query/delete/modify. Add treats recipeIn.recipeID=0 as reserved/invalid and never stores it.
Units: raw REAL values; no scaling. Simultaneous commands are unsupported and modify nothing.
*)

(* CONTRACT_RULES [] *)

tmp_emptyRecipe.recipeID := 0;
tmp_emptyRecipe.ingredientType := 0;
tmp_emptyRecipe.ingredientRatio := 0.0;
tmp_emptyRecipe.productionTemperature := 0.0;

recipeAdded := FALSE;
recipeDeleted := FALSE;
recipeModified := FALSE;
recipeQueryResult := tmp_emptyRecipe;
error := FALSE;
status := 0;

tmp_cmdCount := 0;
IF addRecipe THEN
    tmp_cmdCount := tmp_cmdCount + 1;
END_IF;
IF deleteRecipe THEN
    tmp_cmdCount := tmp_cmdCount + 1;
END_IF;
IF modifyRecipe THEN
    tmp_cmdCount := tmp_cmdCount + 1;
END_IF;
IF queryRecipe THEN
    tmp_cmdCount := tmp_cmdCount + 1;
END_IF;

IF tmp_cmdCount > 1 THEN
    error := TRUE;
    status := 16#8006;
    RETURN;
END_IF;

IF addRecipe THEN
    tmp_found := FALSE;
    tmp_index := 0;
    FOR tmp_i := 1 TO 10 DO
        IF recipe[tmp_i].recipeID = recipeIn.recipeID THEN
            tmp_found := TRUE;
            tmp_index := tmp_i;
            EXIT;
        END_IF;
    END_FOR;

    IF tmp_found THEN
        error := TRUE;
        status := 16#8002;
    ELSE
        tmp_emptyIndex := 0;
        FOR tmp_i := 1 TO 10 DO
            IF recipe[tmp_i].recipeID = 0 THEN
                tmp_emptyIndex := tmp_i;
                EXIT;
            END_IF;
        END_FOR;

        IF tmp_emptyIndex = 0 THEN
            error := TRUE;
            status := 16#8003;
        ELSE
            recipe[tmp_emptyIndex] := recipeIn;
            recipeAdded := TRUE;
            error := FALSE;
            status := 0;
        END_IF;
    END_IF;
END_IF;

IF deleteRecipe THEN
    tmp_found := FALSE;
    tmp_index := 0;
    FOR tmp_i := 1 TO 10 DO
        IF (recipe[tmp_i].recipeID <> 0) AND (recipe[tmp_i].recipeID = recipeIn.recipeID) THEN
            tmp_found := TRUE;
            tmp_index := tmp_i;
            EXIT;
        END_IF;
    END_FOR;

    IF NOT tmp_found THEN
        error := TRUE;
        status := 16#8004;
    ELSE
        recipe[tmp_index] := tmp_emptyRecipe;
        recipeDeleted := TRUE;
        error := FALSE;
        status := 0;
    END_IF;
END_IF;

IF modifyRecipe THEN
    tmp_found := FALSE;
    tmp_index := 0;
    FOR tmp_i := 1 TO 10 DO
        IF (recipe[tmp_i].recipeID <> 0) AND (recipe[tmp_i].recipeID = recipeIn.recipeID) THEN
            tmp_found := TRUE;
            tmp_index := tmp_i;
            EXIT;
        END_IF;
    END_FOR;

    IF NOT tmp_found THEN
        error := TRUE;
        status := 16#8005;
    ELSE
        recipe[tmp_index] := recipeIn;
        recipeModified := TRUE;
        error := FALSE;
        status := 0;
    END_IF;
END_IF;

IF queryRecipe THEN
    tmp_found := FALSE;
    tmp_index := 0;
    FOR tmp_i := 1 TO 10 DO
        IF (recipe[tmp_i].recipeID <> 0) AND (recipe[tmp_i].recipeID = recipeIn.recipeID) THEN
            tmp_found := TRUE;
            tmp_index := tmp_i;
            EXIT;
        END_IF;
    END_FOR;

    IF NOT tmp_found THEN
        error := TRUE;
        status := 16#8001;
    ELSE
        recipeQueryResult := recipe[tmp_index];
        error := FALSE;
        status := 0;
    END_IF;
END_IF;

END_FUNCTION_BLOCK

(* ---- public-hard-04.candidate_01.st ---- *)
(* ENGINEERING_CONTRACT
  PUB001/PUB002: rising edges of enqueue/dequeue are detected by R_TRIG instances each scan.
  PUB003: reset TRUE clears count/head/tail and returns before processing enq/deq requests.
  PUB004: elementCount equals stored count, range 0..capacity; capacity from buffer array length.
  PUB005: rejected full enqueue sets status 16#8002; rejected empty dequeue sets status 16#8001.
  PUB006: first invocation initializes empty state; head/tail/count are internal only.
  PUB007-PUB011: VARIANT buffer/item are accessed via __VARINFO and raw byte copy.
  Unspecified: simultaneous enqueue+dequeue is processed dequeue first, then enqueue.
  Unspecified: invalid buffer metadata leaves the block uninitialized with status 16#0000.
*)
(* CONTRACT_RULES [] *)

TYPE VAR_INFO :
STRUCT
    udiSize : UDINT;
    udiAlignment : UDINT;
    pbyData : POINTER TO BYTE;
    udiTypeClass : UDINT;
    udiTypeSubClass : UDINT;
    udiArrayLength : UDINT;
    sName : STRING(255);
END_STRUCT
END_TYPE;

FUNCTION_BLOCK FB_FIFO
VAR_INPUT
    enqueue : BOOL;
    dequeue : BOOL;
    reset : BOOL;
END_VAR
VAR_OUTPUT
    elementCount : DINT;
    status : WORD;
END_VAR
VAR_IN_OUT
    item : VARIANT;
    buffer : VARIANT;
END_VAR
VAR
    rtEnq : R_TRIG;
    rtDeq : R_TRIG;

    init : BOOL := FALSE;
    capacity : DINT := 0;
    count : DINT := 0;
    head : UDINT := 0;
    tail : UDINT := 0;

    elemSize : UDINT := 0;
    pBuf : POINTER TO BYTE;
    pItem : POINTER TO BYTE;

    infoBuf : VAR_INFO;
    infoItem : VAR_INFO;

    i : UDINT;
    pSrc : POINTER TO BYTE;
    pDst : POINTER TO BYTE;

    tmpEnq : BOOL;
    tmpDeq : BOOL;
END_VAR

rtEnq(CLK := enqueue);
rtDeq(CLK := dequeue);
tmpEnq := rtEnq.Q;
tmpDeq := rtDeq.Q;

elementCount := 0;
status := 16#0000;

IF NOT init THEN
    __VARINFO(ADR(buffer), ADR(infoBuf));
    __VARINFO(ADR(item), ADR(infoItem));

    IF infoBuf.udiArrayLength > 0 THEN
        capacity := TO_DINT(infoBuf.udiArrayLength);
        elemSize := infoItem.udiSize;
        IF elemSize = 0 THEN
            elemSize := 1;
        END_IF;
        pBuf := infoBuf.pbyData;
        pItem := infoItem.pbyData;
        head := 0;
        tail := 0;
        count := 0;
        init := TRUE;
    ELSE
        elementCount := 0;
        status := 16#0000;
        RETURN;
    END_IF;
END_IF;

IF reset THEN
    head := 0;
    tail := 0;
    count := 0;
    elementCount := 0;
    status := 16#0000;
    RETURN;
END_IF;

IF tmpDeq THEN
    IF count > 0 THEN
        pSrc := pBuf + (head * elemSize);
        pDst := pItem;
        FOR i := UDINT#0 TO elemSize - UDINT#1 DO
            pDst[i] := pSrc[i];
        END_FOR;
        head := (head + UDINT#1) MOD TO_UDINT(capacity);
        count := count - 1;
    ELSE
        status := 16#8001;
    END_IF;
END_IF;

IF tmpEnq THEN
    IF count < capacity THEN
        pDst := pBuf + (tail * elemSize);
        pSrc := pItem;
        FOR i := UDINT#0 TO elemSize - UDINT#1 DO
            pDst[i] := pSrc[i];
        END_FOR;
        tail := (tail + UDINT#1) MOD TO_UDINT(capacity);
        count := count + 1;
    ELSE
        IF status = 16#0000 THEN
            status := 16#8002;
        END_IF;
    END_IF;
END_IF;

elementCount := count;

(* ---- public-hard-04.candidate_02.st ---- *)
(* ENGINEERING_CONTRACT
  PUB001/PUB002: rising edges of enqueue/dequeue are detected by R_TRIG instances each scan.
  PUB003: reset TRUE clears count/head/tail and returns before processing enq/deq requests.
  PUB004: elementCount equals stored count, range 0..capacity; capacity from buffer array length.
  PUB005: rejected full enqueue sets status 16#8002; rejected empty dequeue sets status 16#8001.
  PUB006: first invocation initializes empty state; head/tail/count are internal only.
  PUB007-PUB011: VARIANT buffer/item are accessed via __VARINFO and raw byte copy.
  Unspecified: simultaneous enqueue+dequeue is processed dequeue first, then enqueue.
  Unspecified: invalid buffer metadata leaves the block uninitialized with status 16#0000.
*)
(* CONTRACT_RULES [] *)

FUNCTION_BLOCK FB_FIFO
VAR_INPUT
    enqueue : BOOL;
    dequeue : BOOL;
    reset : BOOL;
END_VAR
VAR_OUTPUT
    elementCount : DINT;
    status : WORD;
END_VAR
VAR_IN_OUT
    item : VARIANT;
    buffer : VARIANT;
END_VAR
VAR
    rtEnq : R_TRIG;
    rtDeq : R_TRIG;

    init : BOOL := FALSE;
    capacity : DINT := 0;
    count : DINT := 0;
    head : UDINT := 0;
    tail : UDINT := 0;

    elemSize : UDINT := 0;
    pBuf : POINTER TO BYTE;
    pItem : POINTER TO BYTE;

    infoBuf : __SYSTEM.VAR_INFO;
    infoItem : __SYSTEM.VAR_INFO;

    i : UDINT;
    pSrc : POINTER TO BYTE;
    pDst : POINTER TO BYTE;

    tmpEnq : BOOL;
    tmpDeq : BOOL;
END_VAR

rtEnq(CLK := enqueue);
rtDeq(CLK := dequeue);
tmpEnq := rtEnq.Q;
tmpDeq := rtDeq.Q;

elementCount := 0;
status := 16#0000;

IF NOT init THEN
    __VARINFO(ADR(buffer), ADR(infoBuf));
    __VARINFO(ADR(item), ADR(infoItem));

    IF infoBuf.udiArrayLength > 0 THEN
        capacity := TO_DINT(infoBuf.udiArrayLength);
        elemSize := infoItem.udiSize;
        IF elemSize = 0 THEN
            elemSize := 1;
        END_IF;
        pBuf := infoBuf.pbyData;
        pItem := infoItem.pbyData;
        head := 0;
        tail := 0;
        count := 0;
        init := TRUE;
    ELSE
        elementCount := 0;
        status := 16#0000;
        RETURN;
    END_IF;
END_IF;

IF reset THEN
    head := 0;
    tail := 0;
    count := 0;
    elementCount := 0;
    status := 16#0000;
    RETURN;
END_IF;

IF tmpDeq THEN
    IF count > 0 THEN
        pSrc := pBuf + (head * elemSize);
        pDst := pItem;
        FOR i := UDINT#0 TO elemSize - UDINT#1 DO
            pDst^ := pSrc^;
            pDst := pDst + 1;
            pSrc := pSrc + 1;
        END_FOR;
        head := (head + UDINT#1) MOD TO_UDINT(capacity);
        count := count - 1;
    ELSE
        status := 16#8001;
    END_IF;
END_IF;

IF tmpEnq THEN
    IF count < capacity THEN
        pDst := pBuf + (tail * elemSize);
        pSrc := pItem;
        FOR i := UDINT#0 TO elemSize - UDINT#1 DO
            pDst^ := pSrc^;
            pDst := pDst + 1;
            pSrc := pSrc + 1;
        END_FOR;
        tail := (tail + UDINT#1) MOD TO_UDINT(capacity);
        count := count + 1;
    ELSE
        IF status = 16#0000 THEN
            status := 16#8002;
        END_IF;
    END_IF;
END_IF;

elementCount := count;

END_FUNCTION_BLOCK

(* ---- public-hard-04.candidate_03.st ---- *)
(* ENGINEERING_CONTRACT
  PUB001/PUB002: rising edges of enqueue/dequeue are detected by R_TRIG instances each scan.
  PUB003: reset TRUE clears count/head/tail and returns before processing enq/deq requests.
  PUB004: elementCount equals stored count, range 0..capacity; capacity from buffer array length.
  PUB005: rejected full enqueue sets status 16#8002; rejected empty dequeue sets status 16#8001.
  PUB006: first invocation initializes empty state; head/tail/count are internal only.
  PUB007-PUB011: VARIANT buffer/item are accessed via __VARINFO and raw byte copy.
  Unspecified: simultaneous enqueue+dequeue is processed dequeue first, then enqueue.
  Unspecified: invalid buffer metadata leaves the block uninitialized with status 16#0000.
*)
(* CONTRACT_RULES [] *)

TYPE VAR_INFO :
STRUCT
    udiSize : UDINT;
    udiAlignment : UDINT;
    pbyData : POINTER TO BYTE;
    udiTypeClass : UDINT;
    udiTypeSubClass : UDINT;
    udiArrayLength : UDINT;
    sName : STRING(255);
END_STRUCT
END_TYPE;

FUNCTION_BLOCK FB_FIFO
VAR_INPUT
    enqueue : BOOL;
    dequeue : BOOL;
    reset : BOOL;
END_VAR
VAR_OUTPUT
    elementCount : DINT;
    status : WORD;
END_VAR
VAR_IN_OUT
    item : VARIANT;
    buffer : VARIANT;
END_VAR
VAR
    rtEnq : R_TRIG;
    rtDeq : R_TRIG;

    init : BOOL := FALSE;
    capacity : DINT := 0;
    count : DINT := 0;
    head : UDINT := 0;
    tail : UDINT := 0;

    elemSize : UDINT := 0;
    pBuf : POINTER TO BYTE;
    pItem : POINTER TO BYTE;

    infoBuf : VAR_INFO;
    infoItem : VAR_INFO;

    i : UDINT;
    pSrc : POINTER TO BYTE;
    pDst : POINTER TO BYTE;

    tmpEnq : BOOL;
    tmpDeq : BOOL;
END_VAR

rtEnq(CLK := enqueue);
rtDeq(CLK := dequeue);
tmpEnq := rtEnq.Q;
tmpDeq := rtDeq.Q;

elementCount := 0;
status := 16#0000;

IF NOT init THEN
    __VARINFO(ADR(buffer), ADR(infoBuf));
    __VARINFO(ADR(item), ADR(infoItem));

    IF infoBuf.udiArrayLength > 0 THEN
        capacity := TO_DINT(infoBuf.udiArrayLength);
        elemSize := infoItem.udiSize;
        IF elemSize = 0 THEN
            elemSize := 1;
        END_IF;
        pBuf := infoBuf.pbyData;
        pItem := infoItem.pbyData;
        head := 0;
        tail := 0;
        count := 0;
        init := TRUE;
    ELSE
        elementCount := 0;
        status := 16#0000;
        RETURN;
    END_IF;
END_IF;

IF reset THEN
    head := 0;
    tail := 0;
    count := 0;
    elementCount := 0;
    status := 16#0000;
    RETURN;
END_IF;

IF tmpDeq THEN
    IF count > 0 THEN
        pSrc := pBuf + (head * elemSize);
        pDst := pItem;
        FOR i := UDINT#0 TO (elemSize - UDINT#1) DO
            pDst[i] := pSrc[i];
        END_FOR;
        head := (head + UDINT#1) MOD TO_UDINT(capacity);
        count := count - 1;
    ELSE
        status := 16#8001;
    END_IF;
END_IF;

IF tmpEnq THEN
    IF count < capacity THEN
        pDst := pBuf + (tail * elemSize);
        pSrc := pItem;
        FOR i := UDINT#0 TO (elemSize - UDINT#1) DO
            pDst[i] := pSrc[i];
        END_FOR;
        tail := (tail + UDINT#1) MOD TO_UDINT(capacity);
        count := count + 1;
    ELSE
        IF status = 16#0000 THEN
            status := 16#8002;
        END_IF;
    END_IF;
END_IF;

elementCount := count;
END_FUNCTION_BLOCK

(* ---- public-hard-04.candidate_04.st ---- *)
(* ENGINEERING_CONTRACT
  PUB001/PUB002: rising edges of enqueue/dequeue are detected by R_TRIG instances each scan.
  PUB003: reset TRUE clears count/head/tail and returns before processing enq/deq requests.
  PUB004: elementCount equals stored count, range 0..capacity; capacity from buffer array length.
  PUB005: rejected full enqueue sets status 16#8002; rejected empty dequeue sets status 16#8001.
  PUB006: first invocation initializes empty state; head/tail/count are internal only.
  PUB007-PUB011: VARIANT buffer/item are accessed via __VARINFO and raw byte copy.
  Unspecified: simultaneous enqueue+dequeue is processed dequeue first, then enqueue.
  Unspecified: invalid buffer metadata leaves the block uninitialized with status 16#0000.
*)
(* CONTRACT_RULES [] *)

TYPE VAR_INFO :
STRUCT
    udiSize : UDINT;
    udiAlignment : UDINT;
    pbyData : POINTER TO BYTE;
    udiTypeClass : UDINT;
    udiTypeSubClass : UDINT;
    udiArrayLength : UDINT;
    sName : STRING(255);
END_STRUCT
END_TYPE;

FUNCTION_BLOCK FB_FIFO
VAR_INPUT
    enqueue : BOOL;
    dequeue : BOOL;
    reset : BOOL;
END_VAR
VAR_OUTPUT
    elementCount : DINT;
    status : WORD;
END_VAR
VAR_IN_OUT
    item : VARIANT;
    buffer : VARIANT;
END_VAR
VAR
    rtEnq : R_TRIG;
    rtDeq : R_TRIG;

    init : BOOL := FALSE;
    capacity : DINT := 0;
    count : DINT := 0;
    head : UDINT := 0;
    tail : UDINT := 0;

    elemSize : UDINT := 0;
    pBuf : POINTER TO BYTE;
    pItem : POINTER TO BYTE;

    infoBuf : VAR_INFO;
    infoItem : VAR_INFO;

    i : UDINT;
    pSrc : POINTER TO BYTE;
    pDst : POINTER TO BYTE;

    tmpEnq : BOOL;
    tmpDeq : BOOL;
END_VAR

rtEnq(CLK := enqueue);
rtDeq(CLK := dequeue);
tmpEnq := rtEnq.Q;
tmpDeq := rtDeq.Q;

elementCount := 0;
status := 16#0000;

IF NOT init THEN
    __VARINFO(ADR(buffer), ADR(infoBuf));
    __VARINFO(ADR(item), ADR(infoItem));

    IF infoBuf.udiArrayLength > 0 THEN
        capacity := TO_DINT(infoBuf.udiArrayLength);
        elemSize := infoItem.udiSize;
        IF elemSize = 0 THEN
            elemSize := 1;
        END_IF;
        pBuf := infoBuf.pbyData;
        pItem := infoItem.pbyData;
        head := 0;
        tail := 0;
        count := 0;
        init := TRUE;
    ELSE
        elementCount := 0;
        status := 16#0000;
        RETURN;
    END_IF;
END_IF;

IF reset THEN
    head := 0;
    tail := 0;
    count := 0;
    elementCount := 0;
    status := 16#0000;
    RETURN;
END_IF;

IF tmpDeq THEN
    IF count > 0 THEN
        pSrc := pBuf + (head * elemSize);
        pDst := pItem;
        FOR i := 0 TO elemSize - 1 DO
            pDst[i] := pSrc[i];
        END_FOR;
        head := (head + 1) MOD TO_UDINT(capacity);
        count := count - 1;
    ELSE
        status := 16#8001;
    END_IF;
END_IF;

IF tmpEnq THEN
    IF count < capacity THEN
        pDst := pBuf + (tail * elemSize);
        pSrc := pItem;
        FOR i := 0 TO elemSize - 1 DO
            pDst[i] := pSrc[i];
        END_FOR;
        tail := (tail + 1) MOD TO_UDINT(capacity);
        count := count + 1;
    ELSE
        IF status = 16#0000 THEN
            status := 16#8002;
        END_IF;
    END_IF;
END_IF;

elementCount := count;

END_FUNCTION_BLOCK

(* ---- public-hard-04.raw_candidate_01.st ---- *)
(* ENGINEERING_CONTRACT
  PUB001/PUB002: rising edges of enqueue/dequeue are detected by R_TRIG instances each scan.
  PUB003: reset TRUE clears count/head/tail and returns before processing enq/deq requests.
  PUB004: elementCount equals stored count, range 0..capacity; capacity from buffer array length.
  PUB005: rejected full enqueue sets status 16#8002; rejected empty dequeue sets status 16#8001.
  PUB006: first invocation initializes empty state; head/tail/count are internal only.
  PUB007-PUB011: VARIANT buffer/item are accessed via __VARINFO and raw byte copy.
  Unspecified: simultaneous enqueue+dequeue is processed dequeue first, then enqueue.
  Unspecified: invalid buffer metadata leaves the block uninitialized with status 16#0000.
*)
(* CONTRACT_RULES [] *)

TYPE VAR_INFO :
STRUCT
    udiSize : UDINT;
    udiAlignment : UDINT;
    pbyData : POINTER TO BYTE;
    udiTypeClass : UDINT;
    udiTypeSubClass : UDINT;
    udiArrayLength : UDINT;
    sName : STRING(255);
END_STRUCT
END_TYPE

FUNCTION_BLOCK FB_FIFO
VAR_INPUT
    enqueue : BOOL;
    dequeue : BOOL;
    reset : BOOL;
END_VAR
VAR_OUTPUT
    elementCount : DINT;
    status : WORD;
END_VAR
VAR_IN_OUT
    item : VARIANT;
    buffer : VARIANT;
END_VAR
VAR
    rtEnq : R_TRIG;
    rtDeq : R_TRIG;

    init : BOOL := FALSE;
    capacity : DINT := 0;
    count : DINT := 0;
    head : UDINT := 0;
    tail : UDINT := 0;

    elemSize : UDINT := 0;
    pBuf : POINTER TO BYTE;
    pItem : POINTER TO BYTE;

    infoBuf : VAR_INFO;
    infoItem : VAR_INFO;

    i : UDINT;
    pSrc : POINTER TO BYTE;
    pDst : POINTER TO BYTE;

    tmpEnq : BOOL;
    tmpDeq : BOOL;
END_VAR

rtEnq(CLK := enqueue);
rtDeq(CLK := dequeue);
tmpEnq := rtEnq.Q;
tmpDeq := rtDeq.Q;

elementCount := 0;
status := 16#0000;

IF NOT init THEN
    __VARINFO(ADR(buffer), ADR(infoBuf));
    __VARINFO(ADR(item), ADR(infoItem));

    IF infoBuf.udiArrayLength > 0 THEN
        capacity := TO_DINT(infoBuf.udiArrayLength);
        elemSize := infoItem.udiSize;
        IF elemSize = 0 THEN
            elemSize := 1;
        END_IF
        pBuf := infoBuf.pbyData;
        pItem := infoItem.pbyData;
        head := 0;
        tail := 0;
        count := 0;
        init := TRUE;
    ELSE
        elementCount := 0;
        status := 16#0000;
        RETURN;
    END_IF
END_IF

IF reset THEN
    head := 0;
    tail := 0;
    count := 0;
    elementCount := 0;
    status := 16#0000;
    RETURN;
END_IF

IF tmpDeq THEN
    IF count > 0 THEN
        pSrc := pBuf + (head * elemSize);
        pDst := pItem;
        FOR i := UDINT#0 TO elemSize - UDINT#1 DO
            pDst[i] := pSrc[i];
        END_FOR
        head := (head + UDINT#1) MOD TO_UDINT(capacity);
        count := count - 1;
    ELSE
        status := 16#8001;
    END_IF
END_IF

IF tmpEnq THEN
    IF count < capacity THEN
        pDst := pBuf + (tail * elemSize);
        pSrc := pItem;
        FOR i := UDINT#0 TO elemSize - UDINT#1 DO
            pDst[i] := pSrc[i];
        END_FOR
        tail := (tail + UDINT#1) MOD TO_UDINT(capacity);
        count := count + 1;
    ELSE
        IF status = 16#0000 THEN
            status := 16#8002;
        END_IF
    END_IF
END_IF

elementCount := count;

(* ---- public-hard-04.raw_candidate_02.st ---- *)
(* ENGINEERING_CONTRACT
  PUB001/PUB002: rising edges of enqueue/dequeue are detected by R_TRIG instances each scan.
  PUB003: reset TRUE clears count/head/tail and returns before processing enq/deq requests.
  PUB004: elementCount equals stored count, range 0..capacity; capacity from buffer array length.
  PUB005: rejected full enqueue sets status 16#8002; rejected empty dequeue sets status 16#8001.
  PUB006: first invocation initializes empty state; head/tail/count are internal only.
  PUB007-PUB011: VARIANT buffer/item are accessed via __VARINFO and raw byte copy.
  Unspecified: simultaneous enqueue+dequeue is processed dequeue first, then enqueue.
  Unspecified: invalid buffer metadata leaves the block uninitialized with status 16#0000.
*)
(* CONTRACT_RULES [] *)

FUNCTION_BLOCK FB_FIFO
VAR_INPUT
    enqueue : BOOL;
    dequeue : BOOL;
    reset : BOOL;
END_VAR
VAR_OUTPUT
    elementCount : DINT;
    status : WORD;
END_VAR
VAR_IN_OUT
    item : VARIANT;
    buffer : VARIANT;
END_VAR
VAR
    rtEnq : R_TRIG;
    rtDeq : R_TRIG;

    init : BOOL := FALSE;
    capacity : DINT := 0;
    count : DINT := 0;
    head : UDINT := 0;
    tail : UDINT := 0;

    elemSize : UDINT := 0;
    pBuf : POINTER TO BYTE;
    pItem : POINTER TO BYTE;

    infoBuf : __SYSTEM.VAR_INFO;
    infoItem : __SYSTEM.VAR_INFO;

    i : UDINT;
    pSrc : POINTER TO BYTE;
    pDst : POINTER TO BYTE;

    tmpEnq : BOOL;
    tmpDeq : BOOL;
END_VAR

rtEnq(CLK := enqueue);
rtDeq(CLK := dequeue);
tmpEnq := rtEnq.Q;
tmpDeq := rtDeq.Q;

elementCount := 0;
status := 16#0000;

IF NOT init THEN
    __VARINFO(ADR(buffer), ADR(infoBuf));
    __VARINFO(ADR(item), ADR(infoItem));

    IF infoBuf.udiArrayLength > 0 THEN
        capacity := TO_DINT(infoBuf.udiArrayLength);
        elemSize := infoItem.udiSize;
        IF elemSize = 0 THEN
            elemSize := 1;
        END_IF;
        pBuf := infoBuf.pbyData;
        pItem := infoItem.pbyData;
        head := 0;
        tail := 0;
        count := 0;
        init := TRUE;
    ELSE
        elementCount := 0;
        status := 16#0000;
        RETURN;
    END_IF;
END_IF;

IF reset THEN
    head := 0;
    tail := 0;
    count := 0;
    elementCount := 0;
    status := 16#0000;
    RETURN;
END_IF;

IF tmpDeq THEN
    IF count > 0 THEN
        pSrc := pBuf + (head * elemSize);
        pDst := pItem;
        FOR i := UDINT#0 TO elemSize - UDINT#1 DO
            pDst^ := pSrc^;
            pDst := pDst + 1;
            pSrc := pSrc + 1;
        END_FOR;
        head := (head + UDINT#1) MOD TO_UDINT(capacity);
        count := count - 1;
    ELSE
        status := 16#8001;
    END_IF;
END_IF;

IF tmpEnq THEN
    IF count < capacity THEN
        pDst := pBuf + (tail * elemSize);
        pSrc := pItem;
        FOR i := UDINT#0 TO elemSize - UDINT#1 DO
            pDst^ := pSrc^;
            pDst := pDst + 1;
            pSrc := pSrc + 1;
        END_FOR;
        tail := (tail + UDINT#1) MOD TO_UDINT(capacity);
        count := count + 1;
    ELSE
        IF status = 16#0000 THEN
            status := 16#8002;
        END_IF;
    END_IF;
END_IF;

elementCount := count;

END_FUNCTION_BLOCK

(* ---- public-hard-04.raw_candidate_03.st ---- *)
(* ENGINEERING_CONTRACT
  PUB001/PUB002: rising edges of enqueue/dequeue are detected by R_TRIG instances each scan.
  PUB003: reset TRUE clears count/head/tail and returns before processing enq/deq requests.
  PUB004: elementCount equals stored count, range 0..capacity; capacity from buffer array length.
  PUB005: rejected full enqueue sets status 16#8002; rejected empty dequeue sets status 16#8001.
  PUB006: first invocation initializes empty state; head/tail/count are internal only.
  PUB007-PUB011: VARIANT buffer/item are accessed via __VARINFO and raw byte copy.
  Unspecified: simultaneous enqueue+dequeue is processed dequeue first, then enqueue.
  Unspecified: invalid buffer metadata leaves the block uninitialized with status 16#0000.
*)
(* CONTRACT_RULES [] *)

TYPE VAR_INFO :
STRUCT
    udiSize : UDINT;
    udiAlignment : UDINT;
    pbyData : POINTER TO BYTE;
    udiTypeClass : UDINT;
    udiTypeSubClass : UDINT;
    udiArrayLength : UDINT;
    sName : STRING(255);
END_STRUCT
END_TYPE

FUNCTION_BLOCK FB_FIFO
VAR_INPUT
    enqueue : BOOL;
    dequeue : BOOL;
    reset : BOOL;
END_VAR
VAR_OUTPUT
    elementCount : DINT;
    status : WORD;
END_VAR
VAR_IN_OUT
    item : VARIANT;
    buffer : VARIANT;
END_VAR
VAR
    rtEnq : R_TRIG;
    rtDeq : R_TRIG;

    init : BOOL := FALSE;
    capacity : DINT := 0;
    count : DINT := 0;
    head : UDINT := 0;
    tail : UDINT := 0;

    elemSize : UDINT := 0;
    pBuf : POINTER TO BYTE;
    pItem : POINTER TO BYTE;

    infoBuf : VAR_INFO;
    infoItem : VAR_INFO;

    i : UDINT;
    pSrc : POINTER TO BYTE;
    pDst : POINTER TO BYTE;

    tmpEnq : BOOL;
    tmpDeq : BOOL;
END_VAR

rtEnq(CLK := enqueue);
rtDeq(CLK := dequeue);
tmpEnq := rtEnq.Q;
tmpDeq := rtDeq.Q;

elementCount := 0;
status := 16#0000;

IF NOT init THEN
    __VARINFO(ADR(buffer), ADR(infoBuf));
    __VARINFO(ADR(item), ADR(infoItem));

    IF infoBuf.udiArrayLength > 0 THEN
        capacity := TO_DINT(infoBuf.udiArrayLength);
        elemSize := infoItem.udiSize;
        IF elemSize = 0 THEN
            elemSize := 1;
        END_IF;
        pBuf := infoBuf.pbyData;
        pItem := infoItem.pbyData;
        head := 0;
        tail := 0;
        count := 0;
        init := TRUE;
    ELSE
        elementCount := 0;
        status := 16#0000;
        RETURN;
    END_IF;
END_IF;

IF reset THEN
    head := 0;
    tail := 0;
    count := 0;
    elementCount := 0;
    status := 16#0000;
    RETURN;
END_IF;

IF tmpDeq THEN
    IF count > 0 THEN
        pSrc := pBuf + (head * elemSize);
        pDst := pItem;
        FOR i := UDINT#0 TO (elemSize - UDINT#1) DO
            pDst[i] := pSrc[i];
        END_FOR;
        head := (head + UDINT#1) MOD TO_UDINT(capacity);
        count := count - 1;
    ELSE
        status := 16#8001;
    END_IF;
END_IF;

IF tmpEnq THEN
    IF count < capacity THEN
        pDst := pBuf + (tail * elemSize);
        pSrc := pItem;
        FOR i := UDINT#0 TO (elemSize - UDINT#1) DO
            pDst[i] := pSrc[i];
        END_FOR;
        tail := (tail + UDINT#1) MOD TO_UDINT(capacity);
        count := count + 1;
    ELSE
        IF status = 16#0000 THEN
            status := 16#8002;
        END_IF;
    END_IF;
END_IF;

elementCount := count;
END_FUNCTION_BLOCK

(* ---- public-hard-04.raw_candidate_04.st ---- *)
(* ENGINEERING_CONTRACT
  PUB001/PUB002: rising edges of enqueue/dequeue are detected by R_TRIG instances each scan.
  PUB003: reset TRUE clears count/head/tail and returns before processing enq/deq requests.
  PUB004: elementCount equals stored count, range 0..capacity; capacity from buffer array length.
  PUB005: rejected full enqueue sets status 16#8002; rejected empty dequeue sets status 16#8001.
  PUB006: first invocation initializes empty state; head/tail/count are internal only.
  PUB007-PUB011: VARIANT buffer/item are accessed via __VARINFO and raw byte copy.
  Unspecified: simultaneous enqueue+dequeue is processed dequeue first, then enqueue.
  Unspecified: invalid buffer metadata leaves the block uninitialized with status 16#0000.
*)
(* CONTRACT_RULES [] *)

TYPE VAR_INFO :
STRUCT
    udiSize : UDINT;
    udiAlignment : UDINT;
    pbyData : POINTER TO BYTE;
    udiTypeClass : UDINT;
    udiTypeSubClass : UDINT;
    udiArrayLength : UDINT;
    sName : STRING(255);
END_STRUCT
END_TYPE

FUNCTION_BLOCK FB_FIFO
VAR_INPUT
    enqueue : BOOL;
    dequeue : BOOL;
    reset : BOOL;
END_VAR
VAR_OUTPUT
    elementCount : DINT;
    status : WORD;
END_VAR
VAR_IN_OUT
    item : VARIANT;
    buffer : VARIANT;
END_VAR
VAR
    rtEnq : R_TRIG;
    rtDeq : R_TRIG;

    init : BOOL := FALSE;
    capacity : DINT := 0;
    count : DINT := 0;
    head : UDINT := 0;
    tail : UDINT := 0;

    elemSize : UDINT := 0;
    pBuf : POINTER TO BYTE;
    pItem : POINTER TO BYTE;

    infoBuf : VAR_INFO;
    infoItem : VAR_INFO;

    i : UDINT;
    pSrc : POINTER TO BYTE;
    pDst : POINTER TO BYTE;

    tmpEnq : BOOL;
    tmpDeq : BOOL;
END_VAR

rtEnq(CLK := enqueue);
rtDeq(CLK := dequeue);
tmpEnq := rtEnq.Q;
tmpDeq := rtDeq.Q;

elementCount := 0;
status := 16#0000;

IF NOT init THEN
    __VARINFO(ADR(buffer), ADR(infoBuf));
    __VARINFO(ADR(item), ADR(infoItem));

    IF infoBuf.udiArrayLength > 0 THEN
        capacity := TO_DINT(infoBuf.udiArrayLength);
        elemSize := infoItem.udiSize;
        IF elemSize = 0 THEN
            elemSize := 1;
        END_IF;
        pBuf := infoBuf.pbyData;
        pItem := infoItem.pbyData;
        head := 0;
        tail := 0;
        count := 0;
        init := TRUE;
    ELSE
        elementCount := 0;
        status := 16#0000;
        RETURN;
    END_IF;
END_IF;

IF reset THEN
    head := 0;
    tail := 0;
    count := 0;
    elementCount := 0;
    status := 16#0000;
    RETURN;
END_IF;

IF tmpDeq THEN
    IF count > 0 THEN
        pSrc := pBuf + (head * elemSize);
        pDst := pItem;
        FOR i := 0 TO elemSize - 1 DO
            pDst[i] := pSrc[i];
        END_FOR;
        head := (head + 1) MOD TO_UDINT(capacity);
        count := count - 1;
    ELSE
        status := 16#8001;
    END_IF;
END_IF;

IF tmpEnq THEN
    IF count < capacity THEN
        pDst := pBuf + (tail * elemSize);
        pSrc := pItem;
        FOR i := 0 TO elemSize - 1 DO
            pDst[i] := pSrc[i];
        END_FOR;
        tail := (tail + 1) MOD TO_UDINT(capacity);
        count := count + 1;
    ELSE
        IF status = 16#0000 THEN
            status := 16#8002;
        END_IF;
    END_IF;
END_IF;

elementCount := count;

END_FUNCTION_BLOCK

(* ---- public-hard-05.candidate_01.st ---- *)
FUNCTION_BLOCK MechanicalArmControl
VAR_INPUT
    ManualMode : BOOL;
    SingleStepMode : BOOL;
    SingleCycleMode : BOOL;
    ContinuousMode : BOOL;
    EmergencyStop : BOOL;
    Start : BOOL;
    DownButton : BOOL;
    UpButton : BOOL;
    LeftButton : BOOL;
    RightButton : BOOL;
    GripButton : BOOL;
    ReleaseButton : BOOL;
    DownLimitSwitch : BOOL;
    UpLimitSwitch : BOOL;
    LeftLimitSwitch : BOOL;
    RightLimitSwitch : BOOL;
    GripLimitSwitch : BOOL;
    ReleaseLimitSwitch : BOOL;
END_VAR
VAR_OUTPUT
    MoveDown : BOOL;
    MoveUp : BOOL;
    MoveLeft : BOOL;
    MoveRight : BOOL;
    ActivateGrip : BOOL;
    ActivateRelease : BOOL;
END_VAR
VAR
    local_StartRTrig : R_TRIG;
    local_StartEdge : BOOL;
    local_AutoActive : BOOL := FALSE;
    local_AutoStep : INT := 0;
    local_StepComplete : BOOL;
    local_DesiredMoveDown : BOOL;
    local_DesiredMoveUp : BOOL;
    local_DesiredMoveLeft : BOOL;
    local_DesiredMoveRight : BOOL;
    local_DesiredActivateGrip : BOOL;
    local_DesiredActivateRelease : BOOL;
END_VAR

(* ENGINEERING_CONTRACT
   Manual outputs: active in ManualMode while button=1 and limit=0;
   deactivate on button release, limit reached, or EmergencyStop=FALSE (PUB001, PUB005).
   SingleStep: Start edge begins current step; holds until limit; waits for next Start (PUB002, PUB003).
   SingleCycle: Start edge starts step0; automatic step advance on limit; stops after left (PUB003, PUB015-PUB017).
   Continuous: Start edge starts step0; automatically repeats after left (PUB004, PUB015-PUB017).
   E-stop: all outputs FALSE while EmergencyStop=FALSE; state frozen (PUB005).
   Auto steps 0..7: down,grip,up,right,down,release,up,left; completion via corresponding limit.
   Units/type: BOOL only; no timers; retained state local_AutoActive/local_AutoStep.
*)

(* CONTRACT_RULES [] *)

local_StartRTrig(CLK := Start);
local_StartEdge := local_StartRTrig.Q;

IF NOT EmergencyStop THEN
    MoveDown := FALSE;
    MoveUp := FALSE;
    MoveLeft := FALSE;
    MoveRight := FALSE;
    ActivateGrip := FALSE;
    ActivateRelease := FALSE;
    RETURN;
END_IF;

local_DesiredMoveDown := FALSE;
local_DesiredMoveUp := FALSE;
local_DesiredMoveLeft := FALSE;
local_DesiredMoveRight := FALSE;
local_DesiredActivateGrip := FALSE;
local_DesiredActivateRelease := FALSE;

IF ManualMode THEN
    IF DownButton AND NOT DownLimitSwitch THEN
        local_DesiredMoveDown := TRUE;
    END_IF;
    IF UpButton AND NOT UpLimitSwitch THEN
        local_DesiredMoveUp := TRUE;
    END_IF;
    IF LeftButton AND NOT LeftLimitSwitch THEN
        local_DesiredMoveLeft := TRUE;
    END_IF;
    IF RightButton AND NOT RightLimitSwitch THEN
        local_DesiredMoveRight := TRUE;
    END_IF;
    IF GripButton AND NOT GripLimitSwitch THEN
        local_DesiredActivateGrip := TRUE;
    END_IF;
    IF ReleaseButton AND NOT ReleaseLimitSwitch THEN
        local_DesiredActivateRelease := TRUE;
    END_IF;

ELSIF SingleStepMode OR SingleCycleMode OR ContinuousMode THEN
    IF SingleStepMode THEN
        IF local_StartEdge AND NOT local_AutoActive THEN
            local_AutoActive := TRUE;
        END_IF;

    ELSIF SingleCycleMode THEN
        IF local_StartEdge THEN
            local_AutoStep := 0;
            local_AutoActive := TRUE;
        END_IF;

    ELSIF ContinuousMode THEN
        IF local_StartEdge THEN
            local_AutoStep := 0;
            local_AutoActive := TRUE;
        END_IF;
    END_IF;

    IF local_AutoActive THEN
        CASE local_AutoStep OF
            0: local_DesiredMoveDown := NOT DownLimitSwitch;
            1: local_DesiredActivateGrip := NOT GripLimitSwitch;
            2: local_DesiredMoveUp := NOT UpLimitSwitch;
            3: local_DesiredMoveRight := NOT RightLimitSwitch;
            4: local_DesiredMoveDown := NOT DownLimitSwitch;
            5: local_DesiredActivateRelease := NOT ReleaseLimitSwitch;
            6: local_DesiredMoveUp := NOT UpLimitSwitch;
            7: local_DesiredMoveLeft := NOT LeftLimitSwitch;
        ELSE
            // no active output for invalid step
        END_CASE;
    END_IF;
END_IF;

MoveDown := local_DesiredMoveDown;
MoveUp := local_DesiredMoveUp;
MoveLeft := local_DesiredMoveLeft;
MoveRight := local_DesiredMoveRight;
ActivateGrip := local_DesiredActivateGrip;
ActivateRelease := local_DesiredActivateRelease;

IF SingleStepMode OR SingleCycleMode OR ContinuousMode THEN
    IF local_AutoActive THEN
        local_StepComplete := FALSE;

        IF (local_AutoStep = 0) OR (local_AutoStep = 4) THEN
            local_StepComplete := DownLimitSwitch;
        ELSIF (local_AutoStep = 1) THEN
            local_StepComplete := GripLimitSwitch;
        ELSIF (local_AutoStep = 2) OR (local_AutoStep = 6) THEN
            local_StepComplete := UpLimitSwitch;
        ELSIF (local_AutoStep = 3) THEN
            local_StepComplete := RightLimitSwitch;
        ELSIF (local_AutoStep = 5) THEN
            local_StepComplete := ReleaseLimitSwitch;
        ELSIF (local_AutoStep = 7) THEN
            local_StepComplete := LeftLimitSwitch;
        END_IF;

        IF local_StepComplete THEN
            IF SingleStepMode THEN
                local_AutoActive := FALSE;
                local_AutoStep := (local_AutoStep + 1) MOD 8;

            ELSIF SingleCycleMode THEN
                IF local_AutoStep < 7 THEN
                    local_AutoStep := local_AutoStep + 1;
                    // local_AutoActive remains TRUE
                ELSE
                    local_AutoActive := FALSE;
                    local_AutoStep := 0;
                END_IF;

            ELSIF ContinuousMode THEN
                local_AutoStep := (local_AutoStep + 1) MOD 8;
                local_AutoActive := TRUE;
            END_IF;
        END_IF;
    END_IF;
END_IF;

END_FUNCTION_BLOCK

(* ---- public-hard-05.candidate_02.st ---- *)
FUNCTION_BLOCK MechanicalArmControl
VAR_INPUT
    ManualMode : BOOL;
    SingleStepMode : BOOL;
    SingleCycleMode : BOOL;
    ContinuousMode : BOOL;
    EmergencyStop : BOOL;
    Start : BOOL;
    DownButton : BOOL;
    UpButton : BOOL;
    LeftButton : BOOL;
    RightButton : BOOL;
    GripButton : BOOL;
    ReleaseButton : BOOL;
    DownLimitSwitch : BOOL;
    UpLimitSwitch : BOOL;
    LeftLimitSwitch : BOOL;
    RightLimitSwitch : BOOL;
    GripLimitSwitch : BOOL;
    ReleaseLimitSwitch : BOOL;
END_VAR
VAR_OUTPUT
    MoveDown : BOOL;
    MoveUp : BOOL;
    MoveLeft : BOOL;
    MoveRight : BOOL;
    ActivateGrip : BOOL;
    ActivateRelease : BOOL;
END_VAR
VAR
    local_StartRTrig : R_TRIG;
    local_StartEdge : BOOL;
    local_AutoActive : BOOL := FALSE;
    local_AutoStep : INT := 0;
    local_StepComplete : BOOL;
    local_DesiredMoveDown : BOOL;
    local_DesiredMoveUp : BOOL;
    local_DesiredMoveLeft : BOOL;
    local_DesiredMoveRight : BOOL;
    local_DesiredActivateGrip : BOOL;
    local_DesiredActivateRelease : BOOL;
END_VAR

(* ENGINEERING_CONTRACT
   Manual outputs: active in ManualMode while button=1 and limit=0;
   deactivate on button release, limit reached, or EmergencyStop=FALSE (PUB001, PUB005).
   SingleStep: Start edge begins current step; holds until limit; waits for next Start (PUB002, PUB003).
   SingleCycle: Start edge starts step0; automatic step advance on limit; stops after left (PUB003, PUB015-PUB017).
   Continuous: Start edge starts step0; automatically repeats after left (PUB004, PUB015-PUB017).
   E-stop: all outputs FALSE while EmergencyStop=FALSE; state frozen (PUB005).
   Auto steps 0..7: down,grip,up,right,down,release,up,left; completion via corresponding limit.
   Units/type: BOOL only; no timers; retained state local_AutoActive/local_AutoStep.
*)

(* CONTRACT_RULES [] *)

local_StartRTrig(CLK := Start);
local_StartEdge := local_StartRTrig.Q;

IF NOT EmergencyStop THEN
    MoveDown := FALSE;
    MoveUp := FALSE;
    MoveLeft := FALSE;
    MoveRight := FALSE;
    ActivateGrip := FALSE;
    ActivateRelease := FALSE;
    RETURN;
END_IF;

local_DesiredMoveDown := FALSE;
local_DesiredMoveUp := FALSE;
local_DesiredMoveLeft := FALSE;
local_DesiredMoveRight := FALSE;
local_DesiredActivateGrip := FALSE;
local_DesiredActivateRelease := FALSE;

IF ManualMode THEN
    IF DownButton AND NOT DownLimitSwitch THEN
        local_DesiredMoveDown := TRUE;
    END_IF;
    IF UpButton AND NOT UpLimitSwitch THEN
        local_DesiredMoveUp := TRUE;
    END_IF;
    IF LeftButton AND NOT LeftLimitSwitch THEN
        local_DesiredMoveLeft := TRUE;
    END_IF;
    IF RightButton AND NOT RightLimitSwitch THEN
        local_DesiredMoveRight := TRUE;
    END_IF;
    IF GripButton AND NOT GripLimitSwitch THEN
        local_DesiredActivateGrip := TRUE;
    END_IF;
    IF ReleaseButton AND NOT ReleaseLimitSwitch THEN
        local_DesiredActivateRelease := TRUE;
    END_IF;

ELSIF SingleStepMode OR SingleCycleMode OR ContinuousMode THEN
    IF SingleStepMode THEN
        IF local_StartEdge AND NOT local_AutoActive THEN
            local_AutoActive := TRUE;
        END_IF;

    ELSIF SingleCycleMode THEN
        IF local_StartEdge THEN
            local_AutoStep := 0;
            local_AutoActive := TRUE;
        END_IF;

    ELSIF ContinuousMode THEN
        IF local_StartEdge THEN
            local_AutoStep := 0;
            local_AutoActive := TRUE;
        END_IF;
    END_IF;

    IF local_AutoActive THEN
        CASE local_AutoStep OF
            0: local_DesiredMoveDown := NOT DownLimitSwitch;
            1: local_DesiredActivateGrip := NOT GripLimitSwitch;
            2: local_DesiredMoveUp := NOT UpLimitSwitch;
            3: local_DesiredMoveRight := NOT RightLimitSwitch;
            4: local_DesiredMoveDown := NOT DownLimitSwitch;
            5: local_DesiredActivateRelease := NOT ReleaseLimitSwitch;
            6: local_DesiredMoveUp := NOT UpLimitSwitch;
            7: local_DesiredMoveLeft := NOT LeftLimitSwitch;
        ELSE
            // no active output for invalid step
        END_CASE;
    END_IF;
END_IF;

MoveDown := local_DesiredMoveDown;
MoveUp := local_DesiredMoveUp;
MoveLeft := local_DesiredMoveLeft;
MoveRight := local_DesiredMoveRight;
ActivateGrip := local_DesiredActivateGrip;
ActivateRelease := local_DesiredActivateRelease;

IF SingleStepMode OR SingleCycleMode OR ContinuousMode THEN
    IF local_AutoActive THEN
        local_StepComplete := FALSE;

        IF (local_AutoStep = 0) OR (local_AutoStep = 4) THEN
            local_StepComplete := DownLimitSwitch;
        ELSIF (local_AutoStep = 1) THEN
            local_StepComplete := GripLimitSwitch;
        ELSIF (local_AutoStep = 2) OR (local_AutoStep = 6) THEN
            local_StepComplete := UpLimitSwitch;
        ELSIF (local_AutoStep = 3) THEN
            local_StepComplete := RightLimitSwitch;
        ELSIF (local_AutoStep = 5) THEN
            local_StepComplete := ReleaseLimitSwitch;
        ELSIF (local_AutoStep = 7) THEN
            local_StepComplete := LeftLimitSwitch;
        END_IF;

        IF local_StepComplete THEN
            IF SingleStepMode THEN
                local_AutoActive := FALSE;
                local_AutoStep := (local_AutoStep + 1) MOD 8;

            ELSIF SingleCycleMode THEN
                IF local_AutoStep < 7 THEN
                    local_AutoStep := local_AutoStep + 1;
                    (* local_AutoActive remains TRUE *)
                ELSE
                    local_AutoActive := FALSE;
                    local_AutoStep := 0;
                END_IF;

            ELSIF ContinuousMode THEN
                local_AutoStep := (local_AutoStep + 1) MOD 8;
                local_AutoActive := TRUE;
            END_IF;
        END_IF;
    END_IF;
END_IF;

END_FUNCTION_BLOCK

(* ---- public-hard-05.candidate_03.st ---- *)
FUNCTION_BLOCK MechanicalArmControl
VAR_INPUT
    ManualMode : BOOL;
    SingleStepMode : BOOL;
    SingleCycleMode : BOOL;
    ContinuousMode : BOOL;
    EmergencyStop : BOOL;
    Start : BOOL;
    DownButton : BOOL;
    UpButton : BOOL;
    LeftButton : BOOL;
    RightButton : BOOL;
    GripButton : BOOL;
    ReleaseButton : BOOL;
    DownLimitSwitch : BOOL;
    UpLimitSwitch : BOOL;
    LeftLimitSwitch : BOOL;
    RightLimitSwitch : BOOL;
    GripLimitSwitch : BOOL;
    ReleaseLimitSwitch : BOOL;
END_VAR
VAR_OUTPUT
    MoveDown : BOOL;
    MoveUp : BOOL;
    MoveLeft : BOOL;
    MoveRight : BOOL;
    ActivateGrip : BOOL;
    ActivateRelease : BOOL;
END_VAR
VAR
    local_StartRTrig : R_TRIG;
    local_StartEdge : BOOL;
    local_AutoActive : BOOL := FALSE;
    local_AutoStep : INT := 0;
    local_StepComplete : BOOL;
    local_DesiredMoveDown : BOOL;
    local_DesiredMoveUp : BOOL;
    local_DesiredMoveLeft : BOOL;
    local_DesiredMoveRight : BOOL;
    local_DesiredActivateGrip : BOOL;
    local_DesiredActivateRelease : BOOL;
END_VAR

(* ENGINEERING_CONTRACT
   Manual outputs: active in ManualMode while button=1 and limit=0;
   deactivate on button release, limit reached, or EmergencyStop=FALSE (PUB001, PUB005).
   SingleStep: Start edge begins current step; holds until limit; waits for next Start (PUB002, PUB003).
   SingleCycle: Start edge starts step0; automatic step advance on limit; stops after left (PUB003, PUB015-PUB017).
   Continuous: Start edge starts step0; automatically repeats after left (PUB004, PUB015-PUB017).
   E-stop: all outputs FALSE while EmergencyStop=FALSE; state frozen (PUB005).
   Auto steps 0..7: down,grip,up,right,down,release,up,left; completion via corresponding limit.
   Units/type: BOOL only; no timers; retained state local_AutoActive/local_AutoStep.
*)

(* CONTRACT_RULES [] *)

local_StartRTrig(CLK := Start);
local_StartEdge := local_StartRTrig.Q;

(* Emergency stop has highest priority: immediately clear all outputs and return *)
IF NOT EmergencyStop THEN
    MoveDown := FALSE;
    MoveUp := FALSE;
    MoveLeft := FALSE;
    MoveRight := FALSE;
    ActivateGrip := FALSE;
    ActivateRelease := FALSE;
    RETURN;
END_IF;

(* Initialize desired outputs to FALSE *)
local_DesiredMoveDown := FALSE;
local_DesiredMoveUp := FALSE;
local_DesiredMoveLeft := FALSE;
local_DesiredMoveRight := FALSE;
local_DesiredActivateGrip := FALSE;
local_DesiredActivateRelease := FALSE;

IF ManualMode THEN
    (* Manual control: each action individually driven by its button and limit switch *)
    IF DownButton AND NOT DownLimitSwitch THEN
        local_DesiredMoveDown := TRUE;
    END_IF;
    IF UpButton AND NOT UpLimitSwitch THEN
        local_DesiredMoveUp := TRUE;
    END_IF;
    IF LeftButton AND NOT LeftLimitSwitch THEN
        local_DesiredMoveLeft := TRUE;
    END_IF;
    IF RightButton AND NOT RightLimitSwitch THEN
        local_DesiredMoveRight := TRUE;
    END_IF;
    IF GripButton AND NOT GripLimitSwitch THEN
        local_DesiredActivateGrip := TRUE;
    END_IF;
    IF ReleaseButton AND NOT ReleaseLimitSwitch THEN
        local_DesiredActivateRelease := TRUE;
    END_IF;

ELSIF SingleStepMode OR SingleCycleMode OR ContinuousMode THEN
    (* Automatic modes : single step, single cycle, continuous *)

    IF SingleStepMode THEN
        (* Activate on rising edge of Start only if not already active *)
        IF local_StartEdge AND NOT local_AutoActive THEN
            local_AutoActive := TRUE;
        END_IF;
    ELSIF SingleCycleMode THEN
        (* In single cycle, rising edge of Start resets sequence to step 0 and activates *)
        IF local_StartEdge THEN
            local_AutoStep := 0;
            local_AutoActive := TRUE;
        END_IF;
    ELSIF ContinuousMode THEN
        (* In continuous mode, rising edge of Start resets sequence to step 0 and activates *)
        IF local_StartEdge THEN
            local_AutoStep := 0;
            local_AutoActive := TRUE;
        END_IF;
    END_IF;

    IF local_AutoActive THEN
        CASE local_AutoStep OF
            0: local_DesiredMoveDown := NOT DownLimitSwitch;
            1: local_DesiredActivateGrip := NOT GripLimitSwitch;
            2: local_DesiredMoveUp := NOT UpLimitSwitch;
            3: local_DesiredMoveRight := NOT RightLimitSwitch;
            4: local_DesiredMoveDown := NOT DownLimitSwitch;
            5: local_DesiredActivateRelease := NOT ReleaseLimitSwitch;
            6: local_DesiredMoveUp := NOT UpLimitSwitch;
            7: local_DesiredMoveLeft := NOT LeftLimitSwitch;
        ELSE
            (* Invalid step: no desired movement *)
        END_CASE;
    END_IF;
END_IF;

(* Assign outputs from desired states *)
MoveDown := local_DesiredMoveDown;
MoveUp := local_DesiredMoveUp;
MoveLeft := local_DesiredMoveLeft;
MoveRight := local_DesiredMoveRight;
ActivateGrip := local_DesiredActivateGrip;
ActivateRelease := local_DesiredActivateRelease;

(* Handle step completion and transitions for automatic modes *)
IF SingleStepMode OR SingleCycleMode OR ContinuousMode THEN
    IF local_AutoActive THEN
        local_StepComplete := FALSE;

        IF local_AutoStep = 0 OR local_AutoStep = 4 THEN
            local_StepComplete := DownLimitSwitch;
        ELSIF local_AutoStep = 1 THEN
            local_StepComplete := GripLimitSwitch;
        ELSIF local_AutoStep = 2 OR local_AutoStep = 6 THEN
            local_StepComplete := UpLimitSwitch;
        ELSIF local_AutoStep = 3 THEN
            local_StepComplete := RightLimitSwitch;
        ELSIF local_AutoStep = 5 THEN
            local_StepComplete := ReleaseLimitSwitch;
        ELSIF local_AutoStep = 7 THEN
            local_StepComplete := LeftLimitSwitch;
        END_IF;

        IF local_StepComplete THEN
            IF SingleStepMode THEN
                (* Step finished: deactivate and advance step for next start *)
                local_AutoActive := FALSE;
                local_AutoStep := (local_AutoStep + 1) MOD 8;

            ELSIF SingleCycleMode THEN
                IF local_AutoStep < 7 THEN
                    (* Move to next step in sequence *)
                    local_AutoStep := local_AutoStep + 1;
                    (* local_AutoActive remains TRUE *)
                ELSE
                    (* Cycle complete: stop and reset for next start *)
                    local_AutoActive := FALSE;
                    local_AutoStep := 0;
                END_IF;

            ELSIF ContinuousMode THEN
                (* Automatically advance to next step and continue cycling *)
                local_AutoStep := (local_AutoStep + 1) MOD 8;
                local_AutoActive := TRUE;
            END_IF;
        END_IF;
    END_IF;
END_IF;

END_FUNCTION_BLOCK

(* ---- public-hard-05.candidate_04.st ---- *)
FUNCTION_BLOCK MechanicalArmControl
VAR_INPUT
    ManualMode : BOOL;
    SingleStepMode : BOOL;
    SingleCycleMode : BOOL;
    ContinuousMode : BOOL;
    EmergencyStop : BOOL;
    Start : BOOL;
    DownButton : BOOL;
    UpButton : BOOL;
    LeftButton : BOOL;
    RightButton : BOOL;
    GripButton : BOOL;
    ReleaseButton : BOOL;
    DownLimitSwitch : BOOL;
    UpLimitSwitch : BOOL;
    LeftLimitSwitch : BOOL;
    RightLimitSwitch : BOOL;
    GripLimitSwitch : BOOL;
    ReleaseLimitSwitch : BOOL;
END_VAR
VAR_OUTPUT
    MoveDown : BOOL;
    MoveUp : BOOL;
    MoveLeft : BOOL;
    MoveRight : BOOL;
    ActivateGrip : BOOL;
    ActivateRelease : BOOL;
END_VAR
VAR
    local_StartRTrig : R_TRIG;
    local_StartEdge : BOOL;
    local_AutoActive : BOOL := FALSE;
    local_AutoStep : INT := 0;
    local_StepComplete : BOOL;
    local_DesiredMoveDown : BOOL;
    local_DesiredMoveUp : BOOL;
    local_DesiredMoveLeft : BOOL;
    local_DesiredMoveRight : BOOL;
    local_DesiredActivateGrip : BOOL;
    local_DesiredActivateRelease : BOOL;
END_VAR

(* ENGINEERING_CONTRACT
   Manual outputs: active in ManualMode while button=1 and limit=0;
   deactivate on button release, limit reached, or EmergencyStop=FALSE (PUB001, PUB005).
   SingleStep: Start edge begins current step; holds until limit; waits for next Start (PUB002, PUB003).
   SingleCycle: Start edge starts step0; automatic step advance on limit; stops after left (PUB003, PUB015-PUB017).
   Continuous: Start edge starts step0; automatically repeats after left (PUB004, PUB015-PUB017).
   E-stop: all outputs FALSE while EmergencyStop=FALSE; state frozen (PUB005).
   Auto steps 0..7: down,grip,up,right,down,release,up,left; completion via corresponding limit.
   Units/type: BOOL only; no timers; retained state local_AutoActive/local_AutoStep.
*)

(* CONTRACT_RULES [] *)

local_StartRTrig(CLK := Start);
local_StartEdge := local_StartRTrig.Q;

IF NOT EmergencyStop THEN
    MoveDown := FALSE;
    MoveUp := FALSE;
    MoveLeft := FALSE;
    MoveRight := FALSE;
    ActivateGrip := FALSE;
    ActivateRelease := FALSE;
    RETURN;
END_IF;

local_DesiredMoveDown := FALSE;
local_DesiredMoveUp := FALSE;
local_DesiredMoveLeft := FALSE;
local_DesiredMoveRight := FALSE;
local_DesiredActivateGrip := FALSE;
local_DesiredActivateRelease := FALSE;

IF ManualMode THEN
    IF DownButton AND NOT DownLimitSwitch THEN
        local_DesiredMoveDown := TRUE;
    END_IF;
    IF UpButton AND NOT UpLimitSwitch THEN
        local_DesiredMoveUp := TRUE;
    END_IF;
    IF LeftButton AND NOT LeftLimitSwitch THEN
        local_DesiredMoveLeft := TRUE;
    END_IF;
    IF RightButton AND NOT RightLimitSwitch THEN
        local_DesiredMoveRight := TRUE;
    END_IF;
    IF GripButton AND NOT GripLimitSwitch THEN
        local_DesiredActivateGrip := TRUE;
    END_IF;
    IF ReleaseButton AND NOT ReleaseLimitSwitch THEN
        local_DesiredActivateRelease := TRUE;
    END_IF;

ELSIF SingleStepMode OR SingleCycleMode OR ContinuousMode THEN
    IF SingleStepMode THEN
        IF local_StartEdge AND NOT local_AutoActive THEN
            local_AutoActive := TRUE;
        END_IF;

    ELSIF SingleCycleMode THEN
        IF local_StartEdge THEN
            local_AutoStep := 0;
            local_AutoActive := TRUE;
        END_IF;

    ELSIF ContinuousMode THEN
        IF local_StartEdge THEN
            local_AutoStep := 0;
            local_AutoActive := TRUE;
        END_IF;
    END_IF;

    IF local_AutoActive THEN
        CASE local_AutoStep OF
            0: local_DesiredMoveDown := NOT DownLimitSwitch;
            1: local_DesiredActivateGrip := NOT GripLimitSwitch;
            2: local_DesiredMoveUp := NOT UpLimitSwitch;
            3: local_DesiredMoveRight := NOT RightLimitSwitch;
            4: local_DesiredMoveDown := NOT DownLimitSwitch;
            5: local_DesiredActivateRelease := NOT ReleaseLimitSwitch;
            6: local_DesiredMoveUp := NOT UpLimitSwitch;
            7: local_DesiredMoveLeft := NOT LeftLimitSwitch;
        ELSE
            // no active output for invalid step
        END_CASE;
    END_IF;
END_IF;

MoveDown := local_DesiredMoveDown;
MoveUp := local_DesiredMoveUp;
MoveLeft := local_DesiredMoveLeft;
MoveRight := local_DesiredMoveRight;
ActivateGrip := local_DesiredActivateGrip;
ActivateRelease := local_DesiredActivateRelease;

IF SingleStepMode OR SingleCycleMode OR ContinuousMode THEN
    IF local_AutoActive THEN
        local_StepComplete := FALSE;

        IF (local_AutoStep = 0) OR (local_AutoStep = 4) THEN
            local_StepComplete := DownLimitSwitch;
        ELSIF (local_AutoStep = 1) THEN
            local_StepComplete := GripLimitSwitch;
        ELSIF (local_AutoStep = 2) OR (local_AutoStep = 6) THEN
            local_StepComplete := UpLimitSwitch;
        ELSIF (local_AutoStep = 3) THEN
            local_StepComplete := RightLimitSwitch;
        ELSIF (local_AutoStep = 5) THEN
            local_StepComplete := ReleaseLimitSwitch;
        ELSIF (local_AutoStep = 7) THEN
            local_StepComplete := LeftLimitSwitch;
        END_IF;

        IF local_StepComplete THEN
            IF SingleStepMode THEN
                local_AutoActive := FALSE;
                local_AutoStep := (local_AutoStep + 1) MOD 8;

            ELSIF SingleCycleMode THEN
                IF local_AutoStep < 7 THEN
                    local_AutoStep := local_AutoStep + 1;
                    // local_AutoActive remains TRUE
                ELSE
                    local_AutoActive := FALSE;
                    local_AutoStep := 0;
                END_IF;

            ELSIF ContinuousMode THEN
                local_AutoStep := (local_AutoStep + 1) MOD 8;
                local_AutoActive := TRUE;
            END_IF;
        END_IF;
    END_IF;
END_IF;

END_FUNCTION_BLOCK
